// TIA Portal V19 export
FUNCTION_BLOCK "ALL_VALVES"   // FB1, LAD
{ S7_Optimized_Access := 'TRUE' }
// stored: MemoryReserve 100, SetENOAutomatically false
   VAR
      valve_R1_XV01 { S7_SetPoint := 'True'} : "valve";
      valve_R1_XV02 { S7_SetPoint := 'True'} : "valve";
      valve_R1_XV03 { S7_SetPoint := 'True'} : "valve";
      valve_R1_XV04 { S7_SetPoint := 'True'} : "valve";
      valve_R1_XV05 { S7_SetPoint := 'True'} : "valve";
      valve_R1_XV06 { S7_SetPoint := 'True'} : "valve";
      valve_R1_XV07 { S7_SetPoint := 'True'} : "valve";
      valve_R1_XV08 { S7_SetPoint := 'True'} : "valve";
      valve_R1_XV09 { S7_SetPoint := 'True'} : "valve";
      valve_R1_XV10 { S7_SetPoint := 'True'} : "valve";
      clod_skid { S7_SetPoint := 'True'} : "valve";
      valve_R2_XV01 { S7_SetPoint := 'True'} : "valve";
      valve_R2_XV02 { S7_SetPoint := 'True'} : "valve";
      valve_R2_XV03 { S7_SetPoint := 'True'} : "valve";
      valve_R2_XV04 { S7_SetPoint := 'True'} : "valve";
      valve_R2_XV05 { S7_SetPoint := 'True'} : "valve";
      valve_R2_XV06 { S7_SetPoint := 'True'} : "valve";
      valve_R2_XV07 { S7_SetPoint := 'True'} : "valve";
      valve_R2_XV08 { S7_SetPoint := 'True'} : "valve";
      valve_R2_XV09 { S7_SetPoint := 'True'} : "valve";
      valve_R2_XV10 { S7_SetPoint := 'True'} : "valve";
      valve_R3_XV01 { S7_SetPoint := 'True'} : "valve";
      valve_R3_XV02 { S7_SetPoint := 'True'} : "valve";
      valve_R3_XV03 { S7_SetPoint := 'True'} : "valve";
      valve_R3_XV04 { S7_SetPoint := 'True'} : "valve";
      valve_R3_XV05 { S7_SetPoint := 'True'} : "valve";
      valve_R3_XV06 { S7_SetPoint := 'True'} : "valve";
      valve_R3_XV07 { S7_SetPoint := 'True'} : "valve";
      valve_R3_XV08 { S7_SetPoint := 'True'} : "valve";
      valve_R3_XV09 { S7_SetPoint := 'True'} : "valve";
      valve_R3_XV10 { S7_SetPoint := 'True'} : "valve";
      valve_R4_XV02 { S7_SetPoint := 'True'} : "valve";
      valve_R4_XV01 { S7_SetPoint := 'True'} : "valve";
      valve_R4_XV03 { S7_SetPoint := 'True'} : "valve";
      valve_R4_XV04 { S7_SetPoint := 'True'} : "valve";
      valve_R4_XV05 { S7_SetPoint := 'True'} : "valve";
      valve_R4_XV06 { S7_SetPoint := 'True'} : "valve";
      valve_R4_XV07 { S7_SetPoint := 'True'} : "valve";
      valve_R4_XV08 { S7_SetPoint := 'True'} : "valve";
      valve_R4_XV09 { S7_SetPoint := 'True'} : "valve";
      valve_R4_XV10 { S7_SetPoint := 'True'} : "valve";
      valve_R8_XV2 { S7_SetPoint := 'True'} : "valve";
      valve_R8_XV3 { S7_SetPoint := 'True'} : "valve";
      valve_R8_XV4 { S7_SetPoint := 'True'} : "valve";
      valve_R8_XV5 { S7_SetPoint := 'True'} : "valve";
      valve_R8_XV05 { S7_SetPoint := 'True'} : "valve";
      valve_R8_XV06 { S7_SetPoint := 'True'} : "valve";
      valve_R8_XV07 { S7_SetPoint := 'True'} : "valve";
      valve_R8_XV08 { S7_SetPoint := 'True'} : "valve";
      valve_R8_XV09 { S7_SetPoint := 'True'} : "valve";
      valve_R8_XV10 { S7_SetPoint := 'True'} : "valve";
      valve_R6_XV01 { S7_SetPoint := 'True'} : "valve";
      valve_R6_XV02 { S7_SetPoint := 'True'} : "valve";
      valve_R6_XV03 { S7_SetPoint := 'True'} : "valve";
      valve_R6_XV04 { S7_SetPoint := 'True'} : "valve";
      valve_R6_XV05 { S7_SetPoint := 'True'} : "valve";
      valve_R6_XV06 { S7_SetPoint := 'True'} : "valve";
      valve_R6_XV07 { S7_SetPoint := 'True'} : "valve";
      valve_R6_XV08 { S7_SetPoint := 'True'} : "valve";
      valve_R6_XV09 { S7_SetPoint := 'True'} : "valve";
      valve_R6_XV10 { S7_SetPoint := 'True'} : "valve";
      valve_R7_XV01 { S7_SetPoint := 'True'} : "valve";
      valve_R7_XV02 { S7_SetPoint := 'True'} : "valve";
      valve_R7_XV03 { S7_SetPoint := 'True'} : "valve";
      valve_R7_XV04 { S7_SetPoint := 'True'} : "valve";
      valve_R7_XV05 { S7_SetPoint := 'True'} : "valve";
      valve_R7_XV06 { S7_SetPoint := 'True'} : "valve";
      valve_R7_XV07 { S7_SetPoint := 'True'} : "valve";
      valve_R7_XV08 { S7_SetPoint := 'True'} : "valve";
      valve_R7_XV09 { S7_SetPoint := 'True'} : "valve";
      valve_R7_XV10 { S7_SetPoint := 'True'} : "valve";
      valve_R8_XV01 { S7_SetPoint := 'True'} : "valve";
      valve_R8_XV02 { S7_SetPoint := 'True'} : "valve";
      valve_R8_XV03 { S7_SetPoint := 'True'} : "valve";
      valve_R8_XV04 { S7_SetPoint := 'True'} : "valve";
      valve_R5_XV2 { S7_SetPoint := 'True'} : "valve";
      valve_R5_XV3 { S7_SetPoint := 'True'} : "valve";
      valve_R5_XV4 { S7_SetPoint := 'True'} : "valve";
      valve_R5_XV5 { S7_SetPoint := 'True'} : "valve";
      valve_R5_XV05 { S7_SetPoint := 'True'} : "valve";
      valve_R5_XV06 { S7_SetPoint := 'True'} : "valve";
      valve_R5_XV07 { S7_SetPoint := 'True'} : "valve";
      valve_R5_XV08 { S7_SetPoint := 'True'} : "valve";
      valve_R5_XV09 { S7_SetPoint := 'True'} : "valve";
      valve_R5_XV10 { S7_SetPoint := 'True'} : "valve";
      valve_R9_XV01 { S7_SetPoint := 'True'} : "valve";
      valve_R9_XV02 { S7_SetPoint := 'True'} : "valve";
      valve_R9_XV03 { S7_SetPoint := 'True'} : "valve";
      valve_R9_XV04 { S7_SetPoint := 'True'} : "valve";
      valve_R9_XV05 { S7_SetPoint := 'True'} : "valve";
      valve_R9_XV06 { S7_SetPoint := 'True'} : "valve";
      valve_R9_XV07 { S7_SetPoint := 'True'} : "valve";
      valve_R9_XV08 { S7_SetPoint := 'True'} : "valve";
      valve_R9_XV09 { S7_SetPoint := 'True'} : "valve";
      valve_R9_XV10 { S7_SetPoint := 'True'} : "valve";
      valve_R10_XV01 { S7_SetPoint := 'True'} : "valve";
      valve_R10_XV02 { S7_SetPoint := 'True'} : "valve";
      valve_R10_XV03 { S7_SetPoint := 'True'} : "valve";
      valve_R10_XV04 { S7_SetPoint := 'True'} : "valve";
      valve_R10_XV05 { S7_SetPoint := 'True'} : "valve";
      valve_R10_XV06 { S7_SetPoint := 'True'} : "valve";
      valve_R10_XV07 { S7_SetPoint := 'True'} : "valve";
      valve_R10_XV08 { S7_SetPoint := 'True'} : "valve";
      valve_R10_XV09 { S7_SetPoint := 'True'} : "valve";
      valve_R10_XV10 { S7_SetPoint := 'True'} : "valve";
      valve_R11_XV01 { S7_SetPoint := 'True'} : "valve";
      valve_R11_XV02 { S7_SetPoint := 'True'} : "valve";
      valve_R11_XV03 { S7_SetPoint := 'True'} : "valve";
      valve_R11_XV04 { S7_SetPoint := 'True'} : "valve";
      valve_R11_XV05 { S7_SetPoint := 'True'} : "valve";
      valve_R11_XV06 { S7_SetPoint := 'True'} : "valve";
      valve_R11_XV07 { S7_SetPoint := 'True'} : "valve";
      valve_R11_XV08 { S7_SetPoint := 'True'} : "valve";
      valve_R11_XV09 { S7_SetPoint := 'True'} : "valve";
      valve_R11_XV10 { S7_SetPoint := 'True'} : "valve";
      valve_R12_XV01 { S7_SetPoint := 'True'} : "valve";
      valve_R12_XV02 { S7_SetPoint := 'True'} : "valve";
      valve_R12_XV03 { S7_SetPoint := 'True'} : "valve";
      valve_R12_XV04 { S7_SetPoint := 'True'} : "valve";
      valve_R12_XV05 { S7_SetPoint := 'True'} : "valve";
      valve_R12_XV06 { S7_SetPoint := 'True'} : "valve";
      valve_R12_XV07 { S7_SetPoint := 'True'} : "valve";
      valve_R12_XV08 { S7_SetPoint := 'True'} : "valve";
      valve_R12_XV09 { S7_SetPoint := 'True'} : "valve";
      valve_R12_XV10 { S7_SetPoint := 'True'} : "valve";
      valve_R13_XV01 { S7_SetPoint := 'True'} : "valve";
      valve_R13_XV02 { S7_SetPoint := 'True'} : "valve";
      valve_R13_XV03 { S7_SetPoint := 'True'} : "valve";
      valve_R13_XV04 { S7_SetPoint := 'True'} : "valve";
      valve_R13_XV05 { S7_SetPoint := 'True'} : "valve";
      valve_R13_XV06 { S7_SetPoint := 'True'} : "valve";
      valve_R13_XV07 { S7_SetPoint := 'True'} : "valve";
      valve_R13_XV08 { S7_SetPoint := 'True'} : "valve";
      valve_R13_XV09 { S7_SetPoint := 'True'} : "valve";
      valve_R13_XV10 { S7_SetPoint := 'True'} : "valve";
      valve_R14_XV02 { S7_SetPoint := 'True'} : "valve";
      valve_R14_XV01 { S7_SetPoint := 'True'} : "valve";
      valve_R14_XV03 { S7_SetPoint := 'True'} : "valve";
      valve_R14_XV04 { S7_SetPoint := 'True'} : "valve";
      valve_R14_XV05 { S7_SetPoint := 'True'} : "valve";
      valve_R14_XV06 { S7_SetPoint := 'True'} : "valve";
      valve_R14_XV07 { S7_SetPoint := 'True'} : "valve";
      valve_R14_XV08 { S7_SetPoint := 'True'} : "valve";
      valve_R14_XV09 { S7_SetPoint := 'True'} : "valve";
      valve_R14_XV10 { S7_SetPoint := 'True'} : "valve";
      valve_R15_XV02 { S7_SetPoint := 'True'} : "valve";
      valve_R15_XV01 { S7_SetPoint := 'True'} : "valve";
      valve_R15_XV03 { S7_SetPoint := 'True'} : "valve";
      valve_R15_XV04 { S7_SetPoint := 'True'} : "valve";
      valve_R15_XV05 { S7_SetPoint := 'True'} : "valve";
      valve_R15_XV06 { S7_SetPoint := 'True'} : "valve";
      valve_R15_XV07 { S7_SetPoint := 'True'} : "valve";
      valve_R15_XV08 { S7_SetPoint := 'True'} : "valve";
      valve_R15_XV09 { S7_SetPoint := 'True'} : "valve";
      valve_R15_XV10 { S7_SetPoint := 'True'} : "valve";
      valve_R16_XV02 { S7_SetPoint := 'True'} : "valve";
      valve_R16_XV03 { S7_SetPoint := 'True'} : "valve";
      valve_R16_XV04 { S7_SetPoint := 'True'} : "valve";
      valve_R16_XV05 { S7_SetPoint := 'True'} : "valve";
      valve_R16_XV06 { S7_SetPoint := 'True'} : "valve";
      valve_R16_XV07 { S7_SetPoint := 'True'} : "valve";
      valve_R16_XV08 { S7_SetPoint := 'True'} : "valve";
      valve_R16_XV09 { S7_SetPoint := 'True'} : "valve";
      valve_R16_XV10 { S7_SetPoint := 'True'} : "valve";
      valve_R17_XV01 { S7_SetPoint := 'True'} : "valve";
      valve_R17_XV02 { S7_SetPoint := 'True'} : "valve";
      valve_R17_XV03 { S7_SetPoint := 'True'} : "valve";
      valve_R17_XV04 { S7_SetPoint := 'True'} : "valve";
      valve_R17_XV05 { S7_SetPoint := 'True'} : "valve";
      valve_R17_XV06 { S7_SetPoint := 'True'} : "valve";
      valve_R17_XV07 { S7_SetPoint := 'True'} : "valve";
      valve_R17_XV08 { S7_SetPoint := 'True'} : "valve";
      valve_R17_XV09 { S7_SetPoint := 'True'} : "valve";
      valve_R17_XV10 { S7_SetPoint := 'True'} : "valve";
      valve_R18_XV02 { S7_SetPoint := 'True'} : "valve";
      valve_R18_XV03 { S7_SetPoint := 'True'} : "valve";
      valve_R18_XV04 { S7_SetPoint := 'True'} : "valve";
      valve_R18_XV05 { S7_SetPoint := 'True'} : "valve";
      valve_R18_XV06 { S7_SetPoint := 'True'} : "valve";
      valve_R18_XV07 { S7_SetPoint := 'True'} : "valve";
      valve_R18_XV08 { S7_SetPoint := 'True'} : "valve";
      valve_R18_XV09 { S7_SetPoint := 'True'} : "valve";
      valve_R18_XV10 { S7_SetPoint := 'True'} : "valve";
      child_skid { S7_SetPoint := 'True'} : "valve";
      ultra_child { S7_SetPoint := 'True'} : "valve";
   END_VAR
BEGIN

REGION Network 1: R1_XV01
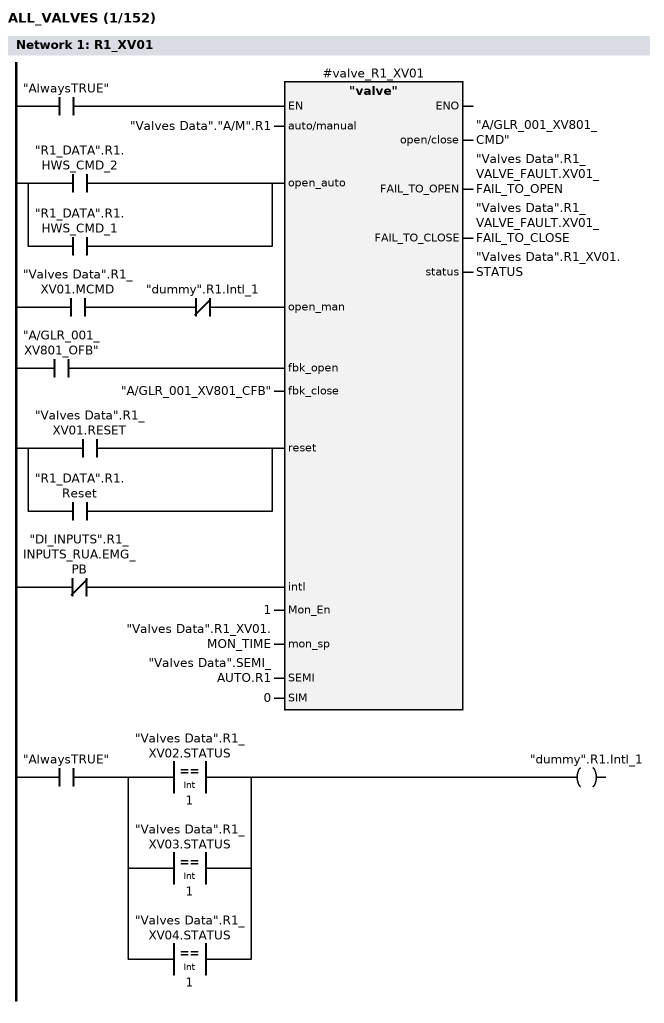
   RUNG wire#powerrail
      Contact( "AlwaysTRUE" )
      #valve_R1_XV01(open_auto := wire#w1, open_man := wire#w2, fbk_open := wire#w3, reset := wire#w4, intl := wire#w5, "auto/manual" := "Valves Data"."A/M".R1, fbk_close := "A/GLR_001_XV801_CFB", Mon_En := 1, mon_sp := "Valves Data".R1_XV01.MON_TIME, SEMI := "Valves Data".SEMI_AUTO.R1, SIM := 0, "open/close" => "A/GLR_001_XV801_CMD", FAIL_TO_OPEN => "Valves Data".R1_VALVE_FAULT.XV01_FAIL_TO_OPEN, FAIL_TO_CLOSE => "Valves Data".R1_VALVE_FAULT.XV01_FAIL_TO_CLOSE, status => "Valves Data".R1_XV01.STATUS)
   END_RUNG
   RUNG wire#powerrail
      Contact( "R1_DATA".R1.HWS_CMD_2 )
   END_RUNG wire#w1
   RUNG wire#powerrail
      Contact( "R1_DATA".R1.HWS_CMD_1 )
   END_RUNG wire#w1
   RUNG wire#powerrail
      Contact( "Valves Data".R1_XV01.MCMD )
      I_Contact( "dummy".R1.Intl_1 )
   END_RUNG wire#w2
   RUNG wire#powerrail
      Contact( "A/GLR_001_XV801_OFB" )
   END_RUNG wire#w3
   RUNG wire#powerrail
      Contact( "Valves Data".R1_XV01.RESET )
   END_RUNG wire#w4
   RUNG wire#powerrail
      Contact( "R1_DATA".R1.Reset )
   END_RUNG wire#w4
   RUNG wire#powerrail
      I_Contact( "DI_INPUTS".R1_INPUTS_RUA.EMG_PB )
   END_RUNG wire#w5
   RUNG wire#powerrail
      Contact( "AlwaysTRUE" )
      wire#w6
      { S7_Templates := "SrcType := Int" } EQ_Contact(in1 := "Valves Data".R1_XV02.STATUS, in2 := 1)
      wire#w7
      Coil( "dummy".R1.Intl_1 )
   END_RUNG
   RUNG wire#w6
      { S7_Templates := "SrcType := Int" } EQ_Contact(in1 := "Valves Data".R1_XV03.STATUS, in2 := 1)
   END_RUNG wire#w7
   RUNG wire#w6
      { S7_Templates := "SrcType := Int" } EQ_Contact(in1 := "Valves Data".R1_XV04.STATUS, in2 := 1)
   END_RUNG wire#w7
   // the same network as SCL:
   IF "AlwaysTRUE" THEN
       #valve_R1_XV01("auto/manual" := "Valves Data"."A/M".R1,   // "valve"
                      open_auto := "R1_DATA".R1.HWS_CMD_2 OR "R1_DATA".R1.HWS_CMD_1,
                      open_man := "Valves Data".R1_XV01.MCMD AND NOT "dummy".R1.Intl_1,
                      fbk_open := "A/GLR_001_XV801_OFB",
                      fbk_close := "A/GLR_001_XV801_CFB",
                      reset := "Valves Data".R1_XV01.RESET OR "R1_DATA".R1.Reset,
                      intl := NOT "DI_INPUTS".R1_INPUTS_RUA.EMG_PB,
                      Mon_En := 1,
                      mon_sp := "Valves Data".R1_XV01.MON_TIME,
                      SEMI := "Valves Data".SEMI_AUTO.R1,
                      SIM := 0,
                      "open/close" => "A/GLR_001_XV801_CMD",
                      FAIL_TO_OPEN => "Valves Data".R1_VALVE_FAULT.XV01_FAIL_TO_OPEN,
                      FAIL_TO_CLOSE => "Valves Data".R1_VALVE_FAULT.XV01_FAIL_TO_CLOSE,
                      status => "Valves Data".R1_XV01.STATUS);
   END_IF;
   "dummy".R1.Intl_1 := "AlwaysTRUE" AND (("Valves Data".R1_XV02.STATUS = 1) OR ("Valves Data".R1_XV03.STATUS = 1) OR ("Valves Data".R1_XV04.STATUS = 1));
END_REGION

REGION Network 2: R1_XV02
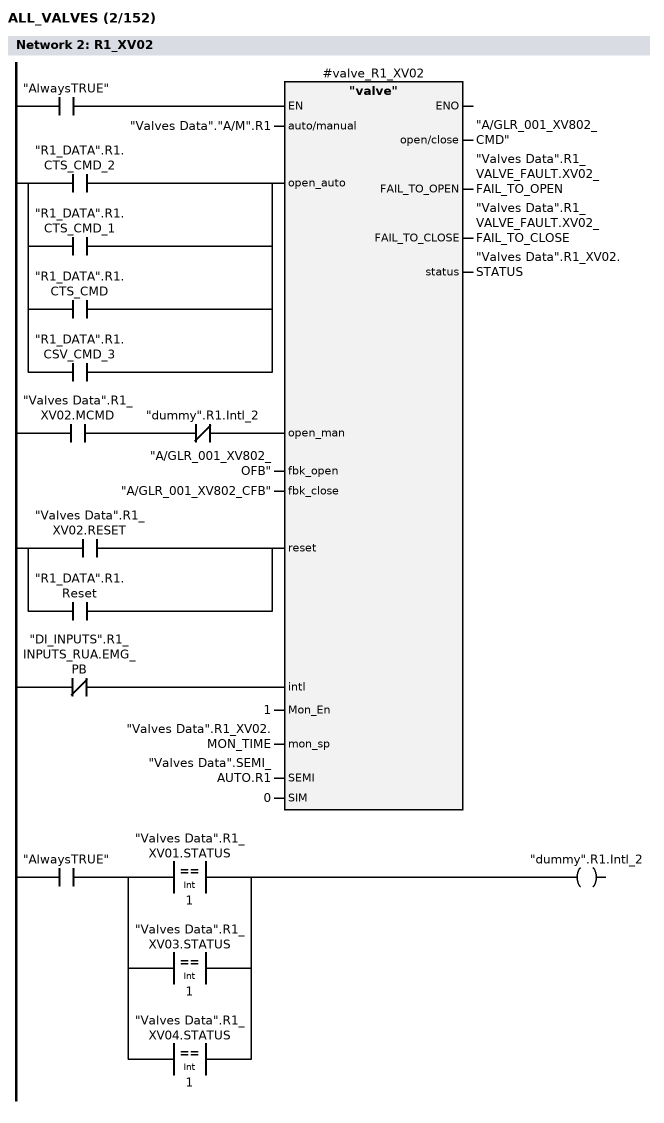
   RUNG wire#powerrail
      Contact( "AlwaysTRUE" )
      #valve_R1_XV02(open_auto := wire#w1, open_man := wire#w2, reset := wire#w3, intl := wire#w4, "auto/manual" := "Valves Data"."A/M".R1, fbk_open := "A/GLR_001_XV802_OFB", fbk_close := "A/GLR_001_XV802_CFB", Mon_En := 1, mon_sp := "Valves Data".R1_XV02.MON_TIME, SEMI := "Valves Data".SEMI_AUTO.R1, SIM := 0, "open/close" => "A/GLR_001_XV802_CMD", FAIL_TO_OPEN => "Valves Data".R1_VALVE_FAULT.XV02_FAIL_TO_OPEN, FAIL_TO_CLOSE => "Valves Data".R1_VALVE_FAULT.XV02_FAIL_TO_CLOSE, status => "Valves Data".R1_XV02.STATUS)
   END_RUNG
   RUNG wire#powerrail
      Contact( "R1_DATA".R1.CTS_CMD_2 )
   END_RUNG wire#w1
   RUNG wire#powerrail
      Contact( "R1_DATA".R1.CTS_CMD_1 )
   END_RUNG wire#w1
   RUNG wire#powerrail
      Contact( "R1_DATA".R1.CTS_CMD )
   END_RUNG wire#w1
   RUNG wire#powerrail
      Contact( "R1_DATA".R1.CSV_CMD_3 )
   END_RUNG wire#w1
   RUNG wire#powerrail
      Contact( "Valves Data".R1_XV02.MCMD )
      I_Contact( "dummy".R1.Intl_2 )
   END_RUNG wire#w2
   RUNG wire#powerrail
      Contact( "Valves Data".R1_XV02.RESET )
   END_RUNG wire#w3
   RUNG wire#powerrail
      Contact( "R1_DATA".R1.Reset )
   END_RUNG wire#w3
   RUNG wire#powerrail
      I_Contact( "DI_INPUTS".R1_INPUTS_RUA.EMG_PB )
   END_RUNG wire#w4
   RUNG wire#powerrail
      Contact( "AlwaysTRUE" )
      wire#w5
      { S7_Templates := "SrcType := Int" } EQ_Contact(in1 := "Valves Data".R1_XV01.STATUS, in2 := 1)
      wire#w6
      Coil( "dummy".R1.Intl_2 )
   END_RUNG
   RUNG wire#w5
      { S7_Templates := "SrcType := Int" } EQ_Contact(in1 := "Valves Data".R1_XV03.STATUS, in2 := 1)
   END_RUNG wire#w6
   RUNG wire#w5
      { S7_Templates := "SrcType := Int" } EQ_Contact(in1 := "Valves Data".R1_XV04.STATUS, in2 := 1)
   END_RUNG wire#w6
   // the same network as SCL:
   IF "AlwaysTRUE" THEN
       #valve_R1_XV02("auto/manual" := "Valves Data"."A/M".R1,   // "valve"
                      open_auto := "R1_DATA".R1.CTS_CMD_2 OR "R1_DATA".R1.CTS_CMD_1 OR "R1_DATA".R1.CTS_CMD OR "R1_DATA".R1.CSV_CMD_3,
                      open_man := "Valves Data".R1_XV02.MCMD AND NOT "dummy".R1.Intl_2,
                      fbk_open := "A/GLR_001_XV802_OFB",
                      fbk_close := "A/GLR_001_XV802_CFB",
                      reset := "Valves Data".R1_XV02.RESET OR "R1_DATA".R1.Reset,
                      intl := NOT "DI_INPUTS".R1_INPUTS_RUA.EMG_PB,
                      Mon_En := 1,
                      mon_sp := "Valves Data".R1_XV02.MON_TIME,
                      SEMI := "Valves Data".SEMI_AUTO.R1,
                      SIM := 0,
                      "open/close" => "A/GLR_001_XV802_CMD",
                      FAIL_TO_OPEN => "Valves Data".R1_VALVE_FAULT.XV02_FAIL_TO_OPEN,
                      FAIL_TO_CLOSE => "Valves Data".R1_VALVE_FAULT.XV02_FAIL_TO_CLOSE,
                      status => "Valves Data".R1_XV02.STATUS);
   END_IF;
   "dummy".R1.Intl_2 := "AlwaysTRUE" AND (("Valves Data".R1_XV01.STATUS = 1) OR ("Valves Data".R1_XV03.STATUS = 1) OR ("Valves Data".R1_XV04.STATUS = 1));
END_REGION

REGION Network 3: R1_XV03
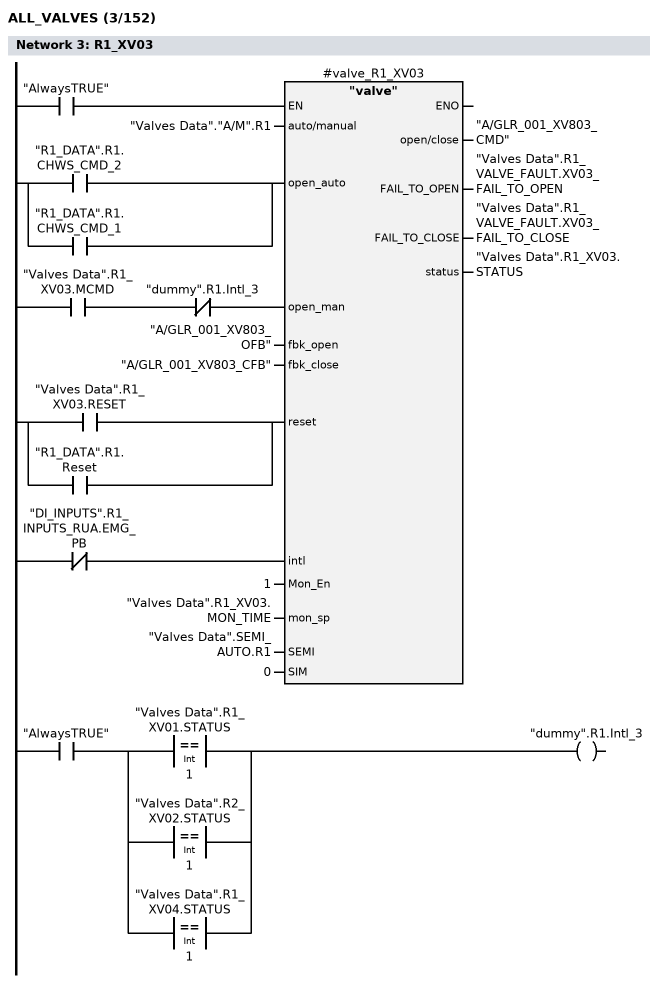
   RUNG wire#powerrail
      Contact( "AlwaysTRUE" )
      #valve_R1_XV03(open_auto := wire#w1, open_man := wire#w2, reset := wire#w3, intl := wire#w4, "auto/manual" := "Valves Data"."A/M".R1, fbk_open := "A/GLR_001_XV803_OFB", fbk_close := "A/GLR_001_XV803_CFB", Mon_En := 1, mon_sp := "Valves Data".R1_XV03.MON_TIME, SEMI := "Valves Data".SEMI_AUTO.R1, SIM := 0, "open/close" => "A/GLR_001_XV803_CMD", FAIL_TO_OPEN => "Valves Data".R1_VALVE_FAULT.XV03_FAIL_TO_OPEN, FAIL_TO_CLOSE => "Valves Data".R1_VALVE_FAULT.XV03_FAIL_TO_CLOSE, status => "Valves Data".R1_XV03.STATUS)
   END_RUNG
   RUNG wire#powerrail
      Contact( "R1_DATA".R1.CHWS_CMD_2 )
   END_RUNG wire#w1
   RUNG wire#powerrail
      Contact( "R1_DATA".R1.CHWS_CMD_1 )
   END_RUNG wire#w1
   RUNG wire#powerrail
      Contact( "Valves Data".R1_XV03.MCMD )
      I_Contact( "dummy".R1.Intl_3 )
   END_RUNG wire#w2
   RUNG wire#powerrail
      Contact( "Valves Data".R1_XV03.RESET )
   END_RUNG wire#w3
   RUNG wire#powerrail
      Contact( "R1_DATA".R1.Reset )
   END_RUNG wire#w3
   RUNG wire#powerrail
      I_Contact( "DI_INPUTS".R1_INPUTS_RUA.EMG_PB )
   END_RUNG wire#w4
   RUNG wire#powerrail
      Contact( "AlwaysTRUE" )
      wire#w5
      { S7_Templates := "SrcType := Int" } EQ_Contact(in1 := "Valves Data".R1_XV01.STATUS, in2 := 1)
      wire#w6
      Coil( "dummy".R1.Intl_3 )
   END_RUNG
   RUNG wire#w5
      { S7_Templates := "SrcType := Int" } EQ_Contact(in1 := "Valves Data".R2_XV02.STATUS, in2 := 1)
   END_RUNG wire#w6
   RUNG wire#w5
      { S7_Templates := "SrcType := Int" } EQ_Contact(in1 := "Valves Data".R1_XV04.STATUS, in2 := 1)
   END_RUNG wire#w6
   // the same network as SCL:
   IF "AlwaysTRUE" THEN
       #valve_R1_XV03("auto/manual" := "Valves Data"."A/M".R1,   // "valve"
                      open_auto := "R1_DATA".R1.CHWS_CMD_2 OR "R1_DATA".R1.CHWS_CMD_1,
                      open_man := "Valves Data".R1_XV03.MCMD AND NOT "dummy".R1.Intl_3,
                      fbk_open := "A/GLR_001_XV803_OFB",
                      fbk_close := "A/GLR_001_XV803_CFB",
                      reset := "Valves Data".R1_XV03.RESET OR "R1_DATA".R1.Reset,
                      intl := NOT "DI_INPUTS".R1_INPUTS_RUA.EMG_PB,
                      Mon_En := 1,
                      mon_sp := "Valves Data".R1_XV03.MON_TIME,
                      SEMI := "Valves Data".SEMI_AUTO.R1,
                      SIM := 0,
                      "open/close" => "A/GLR_001_XV803_CMD",
                      FAIL_TO_OPEN => "Valves Data".R1_VALVE_FAULT.XV03_FAIL_TO_OPEN,
                      FAIL_TO_CLOSE => "Valves Data".R1_VALVE_FAULT.XV03_FAIL_TO_CLOSE,
                      status => "Valves Data".R1_XV03.STATUS);
   END_IF;
   "dummy".R1.Intl_3 := "AlwaysTRUE" AND (("Valves Data".R1_XV01.STATUS = 1) OR ("Valves Data".R2_XV02.STATUS = 1) OR ("Valves Data".R1_XV04.STATUS = 1));
END_REGION

REGION Network 4: R1_XV04
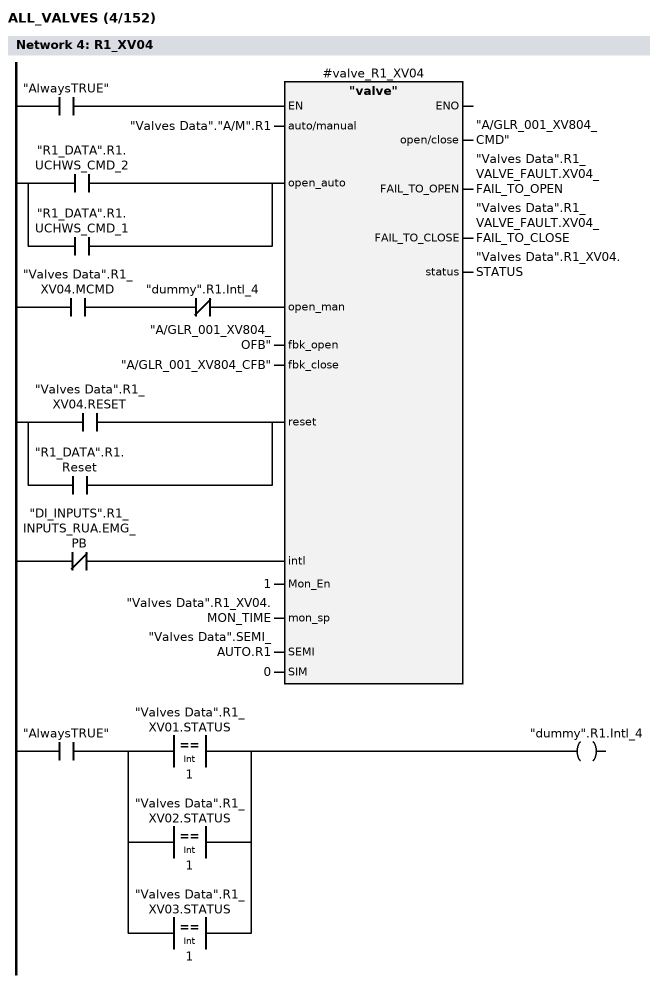
   RUNG wire#powerrail
      Contact( "AlwaysTRUE" )
      #valve_R1_XV04(open_auto := wire#w1, open_man := wire#w2, reset := wire#w3, intl := wire#w4, "auto/manual" := "Valves Data"."A/M".R1, fbk_open := "A/GLR_001_XV804_OFB", fbk_close := "A/GLR_001_XV804_CFB", Mon_En := 1, mon_sp := "Valves Data".R1_XV04.MON_TIME, SEMI := "Valves Data".SEMI_AUTO.R1, SIM := 0, "open/close" => "A/GLR_001_XV804_CMD", FAIL_TO_OPEN => "Valves Data".R1_VALVE_FAULT.XV04_FAIL_TO_OPEN, FAIL_TO_CLOSE => "Valves Data".R1_VALVE_FAULT.XV04_FAIL_TO_CLOSE, status => "Valves Data".R1_XV04.STATUS)
   END_RUNG
   RUNG wire#powerrail
      Contact( "R1_DATA".R1.UCHWS_CMD_2 )
   END_RUNG wire#w1
   RUNG wire#powerrail
      Contact( "R1_DATA".R1.UCHWS_CMD_1 )
   END_RUNG wire#w1
   RUNG wire#powerrail
      Contact( "Valves Data".R1_XV04.MCMD )
      I_Contact( "dummy".R1.Intl_4 )
   END_RUNG wire#w2
   RUNG wire#powerrail
      Contact( "Valves Data".R1_XV04.RESET )
   END_RUNG wire#w3
   RUNG wire#powerrail
      Contact( "R1_DATA".R1.Reset )
   END_RUNG wire#w3
   RUNG wire#powerrail
      I_Contact( "DI_INPUTS".R1_INPUTS_RUA.EMG_PB )
   END_RUNG wire#w4
   RUNG wire#powerrail
      Contact( "AlwaysTRUE" )
      wire#w5
      { S7_Templates := "SrcType := Int" } EQ_Contact(in1 := "Valves Data".R1_XV01.STATUS, in2 := 1)
      wire#w6
      Coil( "dummy".R1.Intl_4 )
   END_RUNG
   RUNG wire#w5
      { S7_Templates := "SrcType := Int" } EQ_Contact(in1 := "Valves Data".R1_XV02.STATUS, in2 := 1)
   END_RUNG wire#w6
   RUNG wire#w5
      { S7_Templates := "SrcType := Int" } EQ_Contact(in1 := "Valves Data".R1_XV03.STATUS, in2 := 1)
   END_RUNG wire#w6
   // the same network as SCL:
   IF "AlwaysTRUE" THEN
       #valve_R1_XV04("auto/manual" := "Valves Data"."A/M".R1,   // "valve"
                      open_auto := "R1_DATA".R1.UCHWS_CMD_2 OR "R1_DATA".R1.UCHWS_CMD_1,
                      open_man := "Valves Data".R1_XV04.MCMD AND NOT "dummy".R1.Intl_4,
                      fbk_open := "A/GLR_001_XV804_OFB",
                      fbk_close := "A/GLR_001_XV804_CFB",
                      reset := "Valves Data".R1_XV04.RESET OR "R1_DATA".R1.Reset,
                      intl := NOT "DI_INPUTS".R1_INPUTS_RUA.EMG_PB,
                      Mon_En := 1,
                      mon_sp := "Valves Data".R1_XV04.MON_TIME,
                      SEMI := "Valves Data".SEMI_AUTO.R1,
                      SIM := 0,
                      "open/close" => "A/GLR_001_XV804_CMD",
                      FAIL_TO_OPEN => "Valves Data".R1_VALVE_FAULT.XV04_FAIL_TO_OPEN,
                      FAIL_TO_CLOSE => "Valves Data".R1_VALVE_FAULT.XV04_FAIL_TO_CLOSE,
                      status => "Valves Data".R1_XV04.STATUS);
   END_IF;
   "dummy".R1.Intl_4 := "AlwaysTRUE" AND (("Valves Data".R1_XV01.STATUS = 1) OR ("Valves Data".R1_XV02.STATUS = 1) OR ("Valves Data".R1_XV03.STATUS = 1));
END_REGION

REGION Network 5: R1_XV05
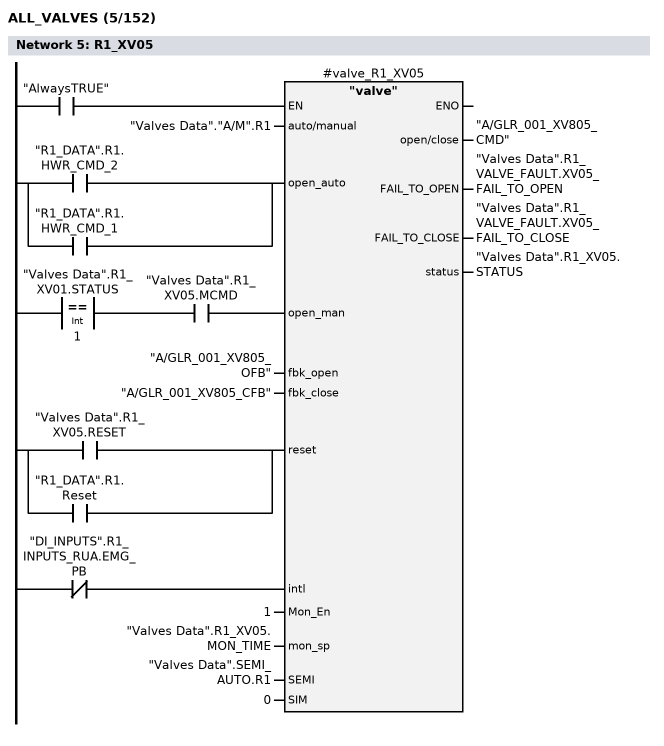
   RUNG wire#powerrail
      Contact( "AlwaysTRUE" )
      #valve_R1_XV05(open_auto := wire#w1, open_man := wire#w2, reset := wire#w3, intl := wire#w4, "auto/manual" := "Valves Data"."A/M".R1, fbk_open := "A/GLR_001_XV805_OFB", fbk_close := "A/GLR_001_XV805_CFB", Mon_En := 1, mon_sp := "Valves Data".R1_XV05.MON_TIME, SEMI := "Valves Data".SEMI_AUTO.R1, SIM := 0, "open/close" => "A/GLR_001_XV805_CMD", FAIL_TO_OPEN => "Valves Data".R1_VALVE_FAULT.XV05_FAIL_TO_OPEN, FAIL_TO_CLOSE => "Valves Data".R1_VALVE_FAULT.XV05_FAIL_TO_CLOSE, status => "Valves Data".R1_XV05.STATUS)
   END_RUNG
   RUNG wire#powerrail
      Contact( "R1_DATA".R1.HWR_CMD_2 )
   END_RUNG wire#w1
   RUNG wire#powerrail
      Contact( "R1_DATA".R1.HWR_CMD_1 )
   END_RUNG wire#w1
   RUNG wire#powerrail
      { S7_Templates := "SrcType := Int" } EQ_Contact(in1 := "Valves Data".R1_XV01.STATUS, in2 := 1)
      Contact( "Valves Data".R1_XV05.MCMD )
   END_RUNG wire#w2
   RUNG wire#powerrail
      Contact( "Valves Data".R1_XV05.RESET )
   END_RUNG wire#w3
   RUNG wire#powerrail
      Contact( "R1_DATA".R1.Reset )
   END_RUNG wire#w3
   RUNG wire#powerrail
      I_Contact( "DI_INPUTS".R1_INPUTS_RUA.EMG_PB )
   END_RUNG wire#w4
   // the same network as SCL:
   IF "AlwaysTRUE" THEN
       #valve_R1_XV05("auto/manual" := "Valves Data"."A/M".R1,   // "valve"
                      open_auto := "R1_DATA".R1.HWR_CMD_2 OR "R1_DATA".R1.HWR_CMD_1,
                      open_man := ("Valves Data".R1_XV01.STATUS = 1) AND "Valves Data".R1_XV05.MCMD,
                      fbk_open := "A/GLR_001_XV805_OFB",
                      fbk_close := "A/GLR_001_XV805_CFB",
                      reset := "Valves Data".R1_XV05.RESET OR "R1_DATA".R1.Reset,
                      intl := NOT "DI_INPUTS".R1_INPUTS_RUA.EMG_PB,
                      Mon_En := 1,
                      mon_sp := "Valves Data".R1_XV05.MON_TIME,
                      SEMI := "Valves Data".SEMI_AUTO.R1,
                      SIM := 0,
                      "open/close" => "A/GLR_001_XV805_CMD",
                      FAIL_TO_OPEN => "Valves Data".R1_VALVE_FAULT.XV05_FAIL_TO_OPEN,
                      FAIL_TO_CLOSE => "Valves Data".R1_VALVE_FAULT.XV05_FAIL_TO_CLOSE,
                      status => "Valves Data".R1_XV05.STATUS);
   END_IF;
END_REGION

REGION Network 6: R1_XV06
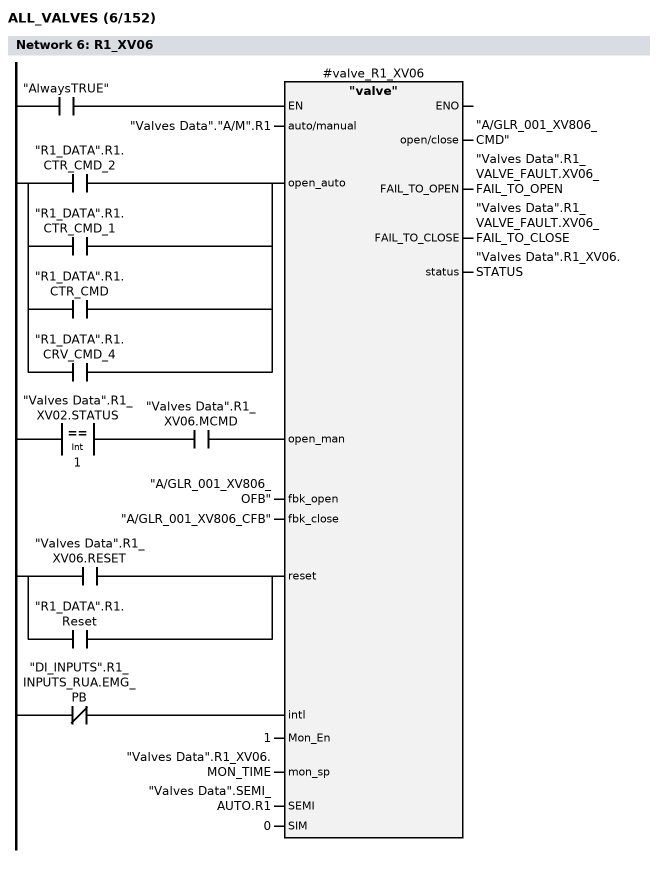
   RUNG wire#powerrail
      Contact( "AlwaysTRUE" )
      #valve_R1_XV06(open_auto := wire#w1, open_man := wire#w2, reset := wire#w3, intl := wire#w4, "auto/manual" := "Valves Data"."A/M".R1, fbk_open := "A/GLR_001_XV806_OFB", fbk_close := "A/GLR_001_XV806_CFB", Mon_En := 1, mon_sp := "Valves Data".R1_XV06.MON_TIME, SEMI := "Valves Data".SEMI_AUTO.R1, SIM := 0, "open/close" => "A/GLR_001_XV806_CMD", FAIL_TO_OPEN => "Valves Data".R1_VALVE_FAULT.XV06_FAIL_TO_OPEN, FAIL_TO_CLOSE => "Valves Data".R1_VALVE_FAULT.XV06_FAIL_TO_CLOSE, status => "Valves Data".R1_XV06.STATUS)
   END_RUNG
   RUNG wire#powerrail
      Contact( "R1_DATA".R1.CTR_CMD_2 )
   END_RUNG wire#w1
   RUNG wire#powerrail
      Contact( "R1_DATA".R1.CTR_CMD_1 )
   END_RUNG wire#w1
   RUNG wire#powerrail
      Contact( "R1_DATA".R1.CTR_CMD )
   END_RUNG wire#w1
   RUNG wire#powerrail
      Contact( "R1_DATA".R1.CRV_CMD_4 )
   END_RUNG wire#w1
   RUNG wire#powerrail
      { S7_Templates := "SrcType := Int" } EQ_Contact(in1 := "Valves Data".R1_XV02.STATUS, in2 := 1)
      Contact( "Valves Data".R1_XV06.MCMD )
   END_RUNG wire#w2
   RUNG wire#powerrail
      Contact( "Valves Data".R1_XV06.RESET )
   END_RUNG wire#w3
   RUNG wire#powerrail
      Contact( "R1_DATA".R1.Reset )
   END_RUNG wire#w3
   RUNG wire#powerrail
      I_Contact( "DI_INPUTS".R1_INPUTS_RUA.EMG_PB )
   END_RUNG wire#w4
   // the same network as SCL:
   IF "AlwaysTRUE" THEN
       #valve_R1_XV06("auto/manual" := "Valves Data"."A/M".R1,   // "valve"
                      open_auto := "R1_DATA".R1.CTR_CMD_2 OR "R1_DATA".R1.CTR_CMD_1 OR "R1_DATA".R1.CTR_CMD OR "R1_DATA".R1.CRV_CMD_4,
                      open_man := ("Valves Data".R1_XV02.STATUS = 1) AND "Valves Data".R1_XV06.MCMD,
                      fbk_open := "A/GLR_001_XV806_OFB",
                      fbk_close := "A/GLR_001_XV806_CFB",
                      reset := "Valves Data".R1_XV06.RESET OR "R1_DATA".R1.Reset,
                      intl := NOT "DI_INPUTS".R1_INPUTS_RUA.EMG_PB,
                      Mon_En := 1,
                      mon_sp := "Valves Data".R1_XV06.MON_TIME,
                      SEMI := "Valves Data".SEMI_AUTO.R1,
                      SIM := 0,
                      "open/close" => "A/GLR_001_XV806_CMD",
                      FAIL_TO_OPEN => "Valves Data".R1_VALVE_FAULT.XV06_FAIL_TO_OPEN,
                      FAIL_TO_CLOSE => "Valves Data".R1_VALVE_FAULT.XV06_FAIL_TO_CLOSE,
                      status => "Valves Data".R1_XV06.STATUS);
   END_IF;
END_REGION

REGION Network 7: R1_XV07
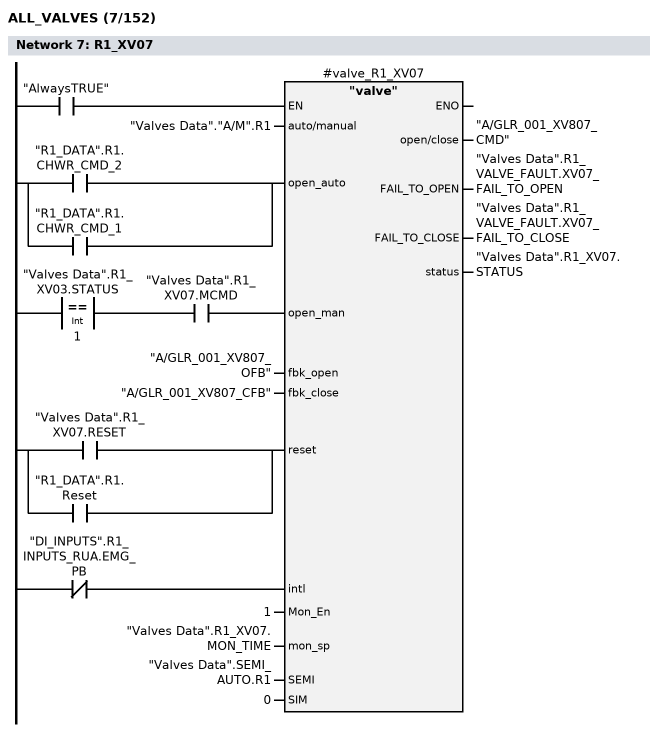
   RUNG wire#powerrail
      Contact( "AlwaysTRUE" )
      #valve_R1_XV07(open_auto := wire#w1, open_man := wire#w2, reset := wire#w3, intl := wire#w4, "auto/manual" := "Valves Data"."A/M".R1, fbk_open := "A/GLR_001_XV807_OFB", fbk_close := "A/GLR_001_XV807_CFB", Mon_En := 1, mon_sp := "Valves Data".R1_XV07.MON_TIME, SEMI := "Valves Data".SEMI_AUTO.R1, SIM := 0, "open/close" => "A/GLR_001_XV807_CMD", FAIL_TO_OPEN => "Valves Data".R1_VALVE_FAULT.XV07_FAIL_TO_OPEN, FAIL_TO_CLOSE => "Valves Data".R1_VALVE_FAULT.XV07_FAIL_TO_CLOSE, status => "Valves Data".R1_XV07.STATUS)
   END_RUNG
   RUNG wire#powerrail
      Contact( "R1_DATA".R1.CHWR_CMD_2 )
   END_RUNG wire#w1
   RUNG wire#powerrail
      Contact( "R1_DATA".R1.CHWR_CMD_1 )
   END_RUNG wire#w1
   RUNG wire#powerrail
      { S7_Templates := "SrcType := Int" } EQ_Contact(in1 := "Valves Data".R1_XV03.STATUS, in2 := 1)
      Contact( "Valves Data".R1_XV07.MCMD )
   END_RUNG wire#w2
   RUNG wire#powerrail
      Contact( "Valves Data".R1_XV07.RESET )
   END_RUNG wire#w3
   RUNG wire#powerrail
      Contact( "R1_DATA".R1.Reset )
   END_RUNG wire#w3
   RUNG wire#powerrail
      I_Contact( "DI_INPUTS".R1_INPUTS_RUA.EMG_PB )
   END_RUNG wire#w4
   // the same network as SCL:
   IF "AlwaysTRUE" THEN
       #valve_R1_XV07("auto/manual" := "Valves Data"."A/M".R1,   // "valve"
                      open_auto := "R1_DATA".R1.CHWR_CMD_2 OR "R1_DATA".R1.CHWR_CMD_1,
                      open_man := ("Valves Data".R1_XV03.STATUS = 1) AND "Valves Data".R1_XV07.MCMD,
                      fbk_open := "A/GLR_001_XV807_OFB",
                      fbk_close := "A/GLR_001_XV807_CFB",
                      reset := "Valves Data".R1_XV07.RESET OR "R1_DATA".R1.Reset,
                      intl := NOT "DI_INPUTS".R1_INPUTS_RUA.EMG_PB,
                      Mon_En := 1,
                      mon_sp := "Valves Data".R1_XV07.MON_TIME,
                      SEMI := "Valves Data".SEMI_AUTO.R1,
                      SIM := 0,
                      "open/close" => "A/GLR_001_XV807_CMD",
                      FAIL_TO_OPEN => "Valves Data".R1_VALVE_FAULT.XV07_FAIL_TO_OPEN,
                      FAIL_TO_CLOSE => "Valves Data".R1_VALVE_FAULT.XV07_FAIL_TO_CLOSE,
                      status => "Valves Data".R1_XV07.STATUS);
   END_IF;
END_REGION

REGION Network 8: R1_XV08
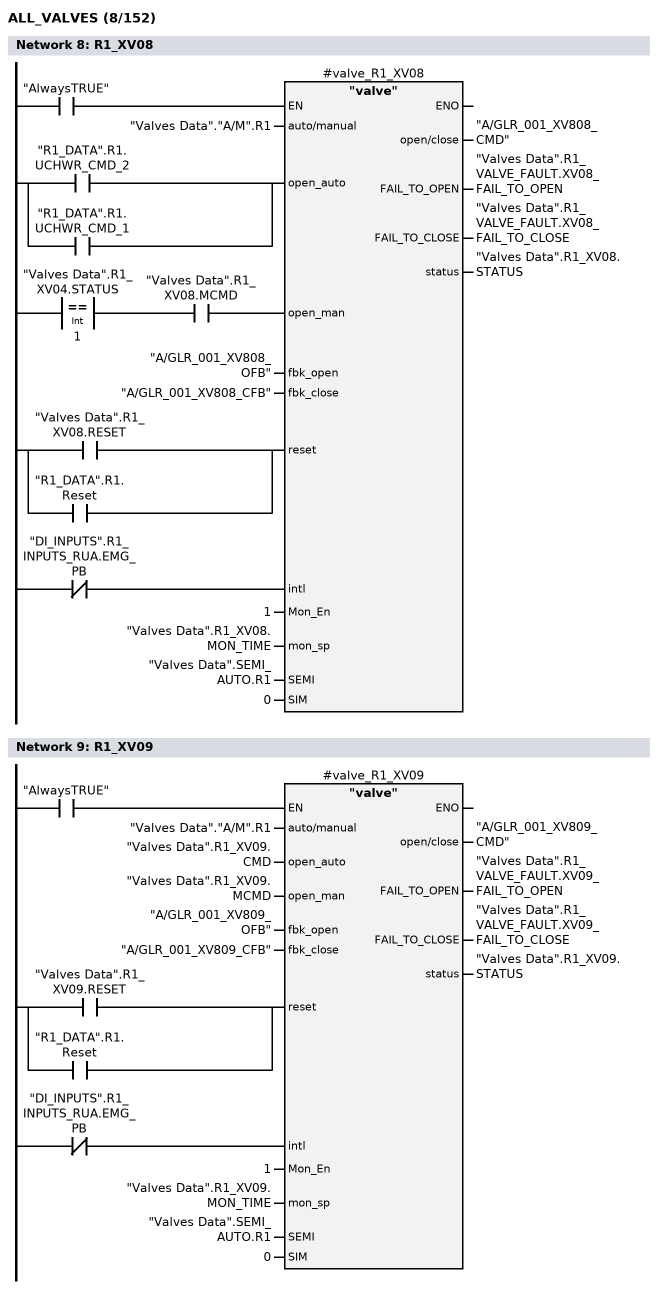
   RUNG wire#powerrail
      Contact( "AlwaysTRUE" )
      #valve_R1_XV08(open_auto := wire#w1, open_man := wire#w2, reset := wire#w3, intl := wire#w4, "auto/manual" := "Valves Data"."A/M".R1, fbk_open := "A/GLR_001_XV808_OFB", fbk_close := "A/GLR_001_XV808_CFB", Mon_En := 1, mon_sp := "Valves Data".R1_XV08.MON_TIME, SEMI := "Valves Data".SEMI_AUTO.R1, SIM := 0, "open/close" => "A/GLR_001_XV808_CMD", FAIL_TO_OPEN => "Valves Data".R1_VALVE_FAULT.XV08_FAIL_TO_OPEN, FAIL_TO_CLOSE => "Valves Data".R1_VALVE_FAULT.XV08_FAIL_TO_CLOSE, status => "Valves Data".R1_XV08.STATUS)
   END_RUNG
   RUNG wire#powerrail
      Contact( "R1_DATA".R1.UCHWR_CMD_2 )
   END_RUNG wire#w1
   RUNG wire#powerrail
      Contact( "R1_DATA".R1.UCHWR_CMD_1 )
   END_RUNG wire#w1
   RUNG wire#powerrail
      { S7_Templates := "SrcType := Int" } EQ_Contact(in1 := "Valves Data".R1_XV04.STATUS, in2 := 1)
      Contact( "Valves Data".R1_XV08.MCMD )
   END_RUNG wire#w2
   RUNG wire#powerrail
      Contact( "Valves Data".R1_XV08.RESET )
   END_RUNG wire#w3
   RUNG wire#powerrail
      Contact( "R1_DATA".R1.Reset )
   END_RUNG wire#w3
   RUNG wire#powerrail
      I_Contact( "DI_INPUTS".R1_INPUTS_RUA.EMG_PB )
   END_RUNG wire#w4
   // the same network as SCL:
   IF "AlwaysTRUE" THEN
       #valve_R1_XV08("auto/manual" := "Valves Data"."A/M".R1,   // "valve"
                      open_auto := "R1_DATA".R1.UCHWR_CMD_2 OR "R1_DATA".R1.UCHWR_CMD_1,
                      open_man := ("Valves Data".R1_XV04.STATUS = 1) AND "Valves Data".R1_XV08.MCMD,
                      fbk_open := "A/GLR_001_XV808_OFB",
                      fbk_close := "A/GLR_001_XV808_CFB",
                      reset := "Valves Data".R1_XV08.RESET OR "R1_DATA".R1.Reset,
                      intl := NOT "DI_INPUTS".R1_INPUTS_RUA.EMG_PB,
                      Mon_En := 1,
                      mon_sp := "Valves Data".R1_XV08.MON_TIME,
                      SEMI := "Valves Data".SEMI_AUTO.R1,
                      SIM := 0,
                      "open/close" => "A/GLR_001_XV808_CMD",
                      FAIL_TO_OPEN => "Valves Data".R1_VALVE_FAULT.XV08_FAIL_TO_OPEN,
                      FAIL_TO_CLOSE => "Valves Data".R1_VALVE_FAULT.XV08_FAIL_TO_CLOSE,
                      status => "Valves Data".R1_XV08.STATUS);
   END_IF;
END_REGION

REGION Network 9: R1_XV09
   RUNG wire#powerrail
      Contact( "AlwaysTRUE" )
      #valve_R1_XV09(reset := wire#w1, intl := wire#w2, "auto/manual" := "Valves Data"."A/M".R1, open_auto := "Valves Data".R1_XV09.CMD, open_man := "Valves Data".R1_XV09.MCMD, fbk_open := "A/GLR_001_XV809_OFB", fbk_close := "A/GLR_001_XV809_CFB", Mon_En := 1, mon_sp := "Valves Data".R1_XV09.MON_TIME, SEMI := "Valves Data".SEMI_AUTO.R1, SIM := 0, "open/close" => "A/GLR_001_XV809_CMD", FAIL_TO_OPEN => "Valves Data".R1_VALVE_FAULT.XV09_FAIL_TO_OPEN, FAIL_TO_CLOSE => "Valves Data".R1_VALVE_FAULT.XV09_FAIL_TO_CLOSE, status => "Valves Data".R1_XV09.STATUS)
   END_RUNG
   RUNG wire#powerrail
      Contact( "Valves Data".R1_XV09.RESET )
   END_RUNG wire#w1
   RUNG wire#powerrail
      Contact( "R1_DATA".R1.Reset )
   END_RUNG wire#w1
   RUNG wire#powerrail
      I_Contact( "DI_INPUTS".R1_INPUTS_RUA.EMG_PB )
   END_RUNG wire#w2
   // the same network as SCL:
   IF "AlwaysTRUE" THEN
       #valve_R1_XV09("auto/manual" := "Valves Data"."A/M".R1,   // "valve"
                      open_auto := "Valves Data".R1_XV09.CMD,
                      open_man := "Valves Data".R1_XV09.MCMD,
                      fbk_open := "A/GLR_001_XV809_OFB",
                      fbk_close := "A/GLR_001_XV809_CFB",
                      reset := "Valves Data".R1_XV09.RESET OR "R1_DATA".R1.Reset,
                      intl := NOT "DI_INPUTS".R1_INPUTS_RUA.EMG_PB,
                      Mon_En := 1,
                      mon_sp := "Valves Data".R1_XV09.MON_TIME,
                      SEMI := "Valves Data".SEMI_AUTO.R1,
                      SIM := 0,
                      "open/close" => "A/GLR_001_XV809_CMD",
                      FAIL_TO_OPEN => "Valves Data".R1_VALVE_FAULT.XV09_FAIL_TO_OPEN,
                      FAIL_TO_CLOSE => "Valves Data".R1_VALVE_FAULT.XV09_FAIL_TO_CLOSE,
                      status => "Valves Data".R1_XV09.STATUS);
   END_IF;
END_REGION

REGION Network 10: R1_XV10
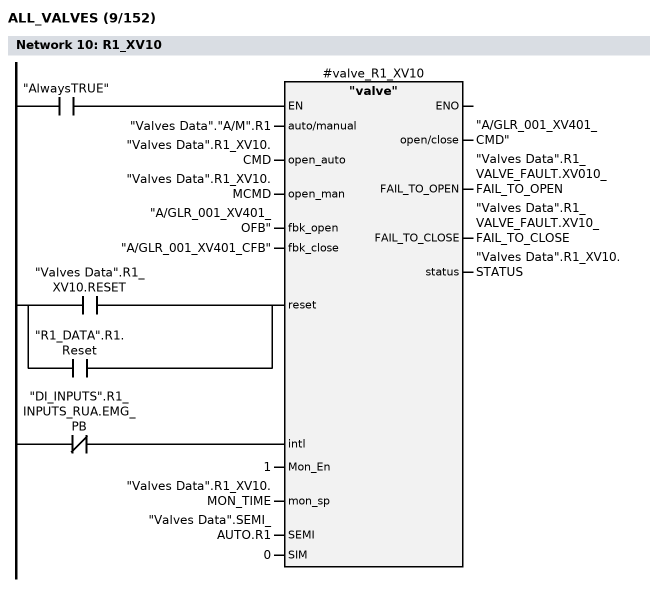
   RUNG wire#powerrail
      Contact( "AlwaysTRUE" )
      #valve_R1_XV10(reset := wire#w1, intl := wire#w2, "auto/manual" := "Valves Data"."A/M".R1, open_auto := "Valves Data".R1_XV10.CMD, open_man := "Valves Data".R1_XV10.MCMD, fbk_open := "A/GLR_001_XV401_OFB", fbk_close := "A/GLR_001_XV401_CFB", Mon_En := 1, mon_sp := "Valves Data".R1_XV10.MON_TIME, SEMI := "Valves Data".SEMI_AUTO.R1, SIM := 0, "open/close" => "A/GLR_001_XV401_CMD", FAIL_TO_OPEN => "Valves Data".R1_VALVE_FAULT.XV010_FAIL_TO_OPEN, FAIL_TO_CLOSE => "Valves Data".R1_VALVE_FAULT.XV10_FAIL_TO_CLOSE, status => "Valves Data".R1_XV10.STATUS)
   END_RUNG
   RUNG wire#powerrail
      Contact( "Valves Data".R1_XV10.RESET )
   END_RUNG wire#w1
   RUNG wire#powerrail
      Contact( "R1_DATA".R1.Reset )
   END_RUNG wire#w1
   RUNG wire#powerrail
      I_Contact( "DI_INPUTS".R1_INPUTS_RUA.EMG_PB )
   END_RUNG wire#w2
   // the same network as SCL:
   IF "AlwaysTRUE" THEN
       #valve_R1_XV10("auto/manual" := "Valves Data"."A/M".R1,   // "valve"
                      open_auto := "Valves Data".R1_XV10.CMD,
                      open_man := "Valves Data".R1_XV10.MCMD,
                      fbk_open := "A/GLR_001_XV401_OFB",
                      fbk_close := "A/GLR_001_XV401_CFB",
                      reset := "Valves Data".R1_XV10.RESET OR "R1_DATA".R1.Reset,
                      intl := NOT "DI_INPUTS".R1_INPUTS_RUA.EMG_PB,
                      Mon_En := 1,
                      mon_sp := "Valves Data".R1_XV10.MON_TIME,
                      SEMI := "Valves Data".SEMI_AUTO.R1,
                      SIM := 0,
                      "open/close" => "A/GLR_001_XV401_CMD",
                      FAIL_TO_OPEN => "Valves Data".R1_VALVE_FAULT.XV010_FAIL_TO_OPEN,
                      FAIL_TO_CLOSE => "Valves Data".R1_VALVE_FAULT.XV10_FAIL_TO_CLOSE,
                      status => "Valves Data".R1_XV10.STATUS);
   END_IF;
END_REGION

REGION Network 11: ****REACTOR_02****
END_REGION

REGION Network 12: R2_XV01
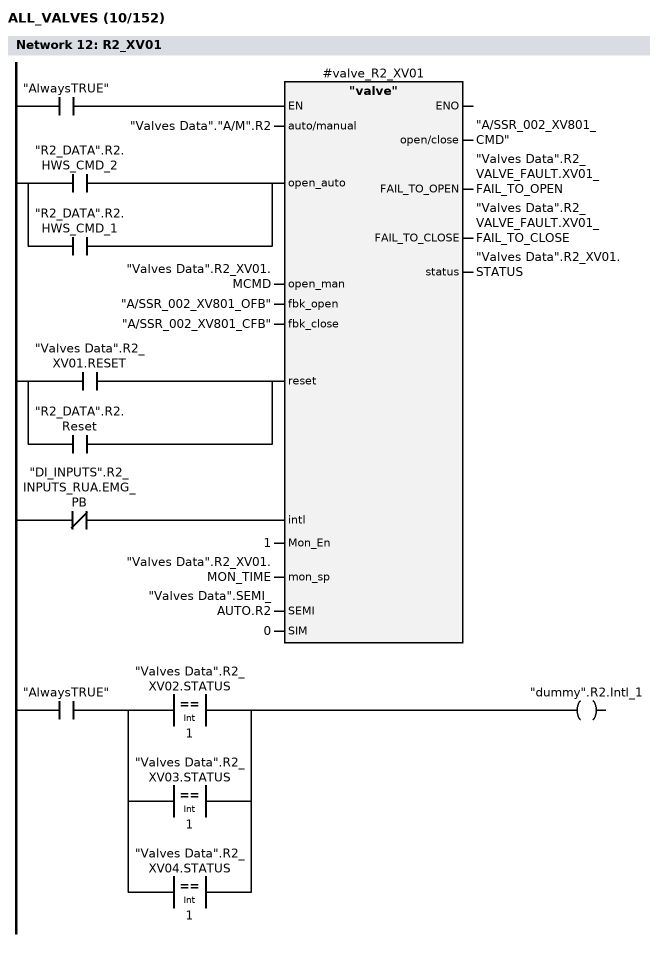
   RUNG wire#powerrail
      Contact( "AlwaysTRUE" )
      #valve_R2_XV01(open_auto := wire#w1, reset := wire#w2, intl := wire#w3, "auto/manual" := "Valves Data"."A/M".R2, open_man := "Valves Data".R2_XV01.MCMD, fbk_open := "A/SSR_002_XV801_OFB", fbk_close := "A/SSR_002_XV801_CFB", Mon_En := 1, mon_sp := "Valves Data".R2_XV01.MON_TIME, SEMI := "Valves Data".SEMI_AUTO.R2, SIM := 0, "open/close" => "A/SSR_002_XV801_CMD", FAIL_TO_OPEN => "Valves Data".R2_VALVE_FAULT.XV01_FAIL_TO_OPEN, FAIL_TO_CLOSE => "Valves Data".R2_VALVE_FAULT.XV01_FAIL_TO_CLOSE, status => "Valves Data".R2_XV01.STATUS)
   END_RUNG
   RUNG wire#powerrail
      Contact( "R2_DATA".R2.HWS_CMD_2 )
   END_RUNG wire#w1
   RUNG wire#powerrail
      Contact( "R2_DATA".R2.HWS_CMD_1 )
   END_RUNG wire#w1
   RUNG wire#powerrail
      Contact( "Valves Data".R2_XV01.RESET )
   END_RUNG wire#w2
   RUNG wire#powerrail
      Contact( "R2_DATA".R2.Reset )
   END_RUNG wire#w2
   RUNG wire#powerrail
      I_Contact( "DI_INPUTS".R2_INPUTS_RUA.EMG_PB )
   END_RUNG wire#w3
   RUNG wire#powerrail
      Contact( "AlwaysTRUE" )
      wire#w4
      { S7_Templates := "SrcType := Int" } EQ_Contact(in1 := "Valves Data".R2_XV02.STATUS, in2 := 1)
      wire#w5
      Coil( "dummy".R2.Intl_1 )
   END_RUNG
   RUNG wire#w4
      { S7_Templates := "SrcType := Int" } EQ_Contact(in1 := "Valves Data".R2_XV03.STATUS, in2 := 1)
   END_RUNG wire#w5
   RUNG wire#w4
      { S7_Templates := "SrcType := Int" } EQ_Contact(in1 := "Valves Data".R2_XV04.STATUS, in2 := 1)
   END_RUNG wire#w5
   // the same network as SCL:
   IF "AlwaysTRUE" THEN
       #valve_R2_XV01("auto/manual" := "Valves Data"."A/M".R2,   // "valve"
                      open_auto := "R2_DATA".R2.HWS_CMD_2 OR "R2_DATA".R2.HWS_CMD_1,
                      open_man := "Valves Data".R2_XV01.MCMD,
                      fbk_open := "A/SSR_002_XV801_OFB",
                      fbk_close := "A/SSR_002_XV801_CFB",
                      reset := "Valves Data".R2_XV01.RESET OR "R2_DATA".R2.Reset,
                      intl := NOT "DI_INPUTS".R2_INPUTS_RUA.EMG_PB,
                      Mon_En := 1,
                      mon_sp := "Valves Data".R2_XV01.MON_TIME,
                      SEMI := "Valves Data".SEMI_AUTO.R2,
                      SIM := 0,
                      "open/close" => "A/SSR_002_XV801_CMD",
                      FAIL_TO_OPEN => "Valves Data".R2_VALVE_FAULT.XV01_FAIL_TO_OPEN,
                      FAIL_TO_CLOSE => "Valves Data".R2_VALVE_FAULT.XV01_FAIL_TO_CLOSE,
                      status => "Valves Data".R2_XV01.STATUS);
   END_IF;
   "dummy".R2.Intl_1 := "AlwaysTRUE" AND (("Valves Data".R2_XV02.STATUS = 1) OR ("Valves Data".R2_XV03.STATUS = 1) OR ("Valves Data".R2_XV04.STATUS = 1));
END_REGION

REGION Network 13: R2_XV02
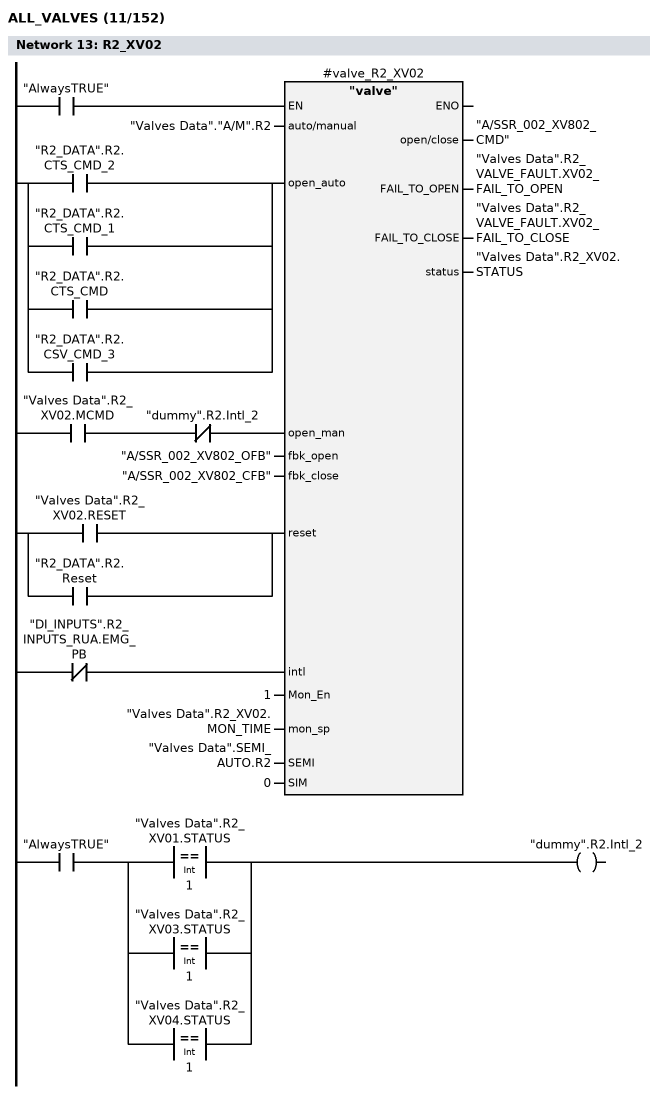
   RUNG wire#powerrail
      Contact( "AlwaysTRUE" )
      #valve_R2_XV02(open_auto := wire#w1, open_man := wire#w2, reset := wire#w3, intl := wire#w4, "auto/manual" := "Valves Data"."A/M".R2, fbk_open := "A/SSR_002_XV802_OFB", fbk_close := "A/SSR_002_XV802_CFB", Mon_En := 1, mon_sp := "Valves Data".R2_XV02.MON_TIME, SEMI := "Valves Data".SEMI_AUTO.R2, SIM := 0, "open/close" => "A/SSR_002_XV802_CMD", FAIL_TO_OPEN => "Valves Data".R2_VALVE_FAULT.XV02_FAIL_TO_OPEN, FAIL_TO_CLOSE => "Valves Data".R2_VALVE_FAULT.XV02_FAIL_TO_CLOSE, status => "Valves Data".R2_XV02.STATUS)
   END_RUNG
   RUNG wire#powerrail
      Contact( "R2_DATA".R2.CTS_CMD_2 )
   END_RUNG wire#w1
   RUNG wire#powerrail
      Contact( "R2_DATA".R2.CTS_CMD_1 )
   END_RUNG wire#w1
   RUNG wire#powerrail
      Contact( "R2_DATA".R2.CTS_CMD )
   END_RUNG wire#w1
   RUNG wire#powerrail
      Contact( "R2_DATA".R2.CSV_CMD_3 )
   END_RUNG wire#w1
   RUNG wire#powerrail
      Contact( "Valves Data".R2_XV02.MCMD )
      I_Contact( "dummy".R2.Intl_2 )
   END_RUNG wire#w2
   RUNG wire#powerrail
      Contact( "Valves Data".R2_XV02.RESET )
   END_RUNG wire#w3
   RUNG wire#powerrail
      Contact( "R2_DATA".R2.Reset )
   END_RUNG wire#w3
   RUNG wire#powerrail
      I_Contact( "DI_INPUTS".R2_INPUTS_RUA.EMG_PB )
   END_RUNG wire#w4
   RUNG wire#powerrail
      Contact( "AlwaysTRUE" )
      wire#w5
      { S7_Templates := "SrcType := Int" } EQ_Contact(in1 := "Valves Data".R2_XV01.STATUS, in2 := 1)
      wire#w6
      Coil( "dummy".R2.Intl_2 )
   END_RUNG
   RUNG wire#w5
      { S7_Templates := "SrcType := Int" } EQ_Contact(in1 := "Valves Data".R2_XV03.STATUS, in2 := 1)
   END_RUNG wire#w6
   RUNG wire#w5
      { S7_Templates := "SrcType := Int" } EQ_Contact(in1 := "Valves Data".R2_XV04.STATUS, in2 := 1)
   END_RUNG wire#w6
   // the same network as SCL:
   IF "AlwaysTRUE" THEN
       #valve_R2_XV02("auto/manual" := "Valves Data"."A/M".R2,   // "valve"
                      open_auto := "R2_DATA".R2.CTS_CMD_2 OR "R2_DATA".R2.CTS_CMD_1 OR "R2_DATA".R2.CTS_CMD OR "R2_DATA".R2.CSV_CMD_3,
                      open_man := "Valves Data".R2_XV02.MCMD AND NOT "dummy".R2.Intl_2,
                      fbk_open := "A/SSR_002_XV802_OFB",
                      fbk_close := "A/SSR_002_XV802_CFB",
                      reset := "Valves Data".R2_XV02.RESET OR "R2_DATA".R2.Reset,
                      intl := NOT "DI_INPUTS".R2_INPUTS_RUA.EMG_PB,
                      Mon_En := 1,
                      mon_sp := "Valves Data".R2_XV02.MON_TIME,
                      SEMI := "Valves Data".SEMI_AUTO.R2,
                      SIM := 0,
                      "open/close" => "A/SSR_002_XV802_CMD",
                      FAIL_TO_OPEN => "Valves Data".R2_VALVE_FAULT.XV02_FAIL_TO_OPEN,
                      FAIL_TO_CLOSE => "Valves Data".R2_VALVE_FAULT.XV02_FAIL_TO_CLOSE,
                      status => "Valves Data".R2_XV02.STATUS);
   END_IF;
   "dummy".R2.Intl_2 := "AlwaysTRUE" AND (("Valves Data".R2_XV01.STATUS = 1) OR ("Valves Data".R2_XV03.STATUS = 1) OR ("Valves Data".R2_XV04.STATUS = 1));
END_REGION

REGION Network 14: R2_XV03
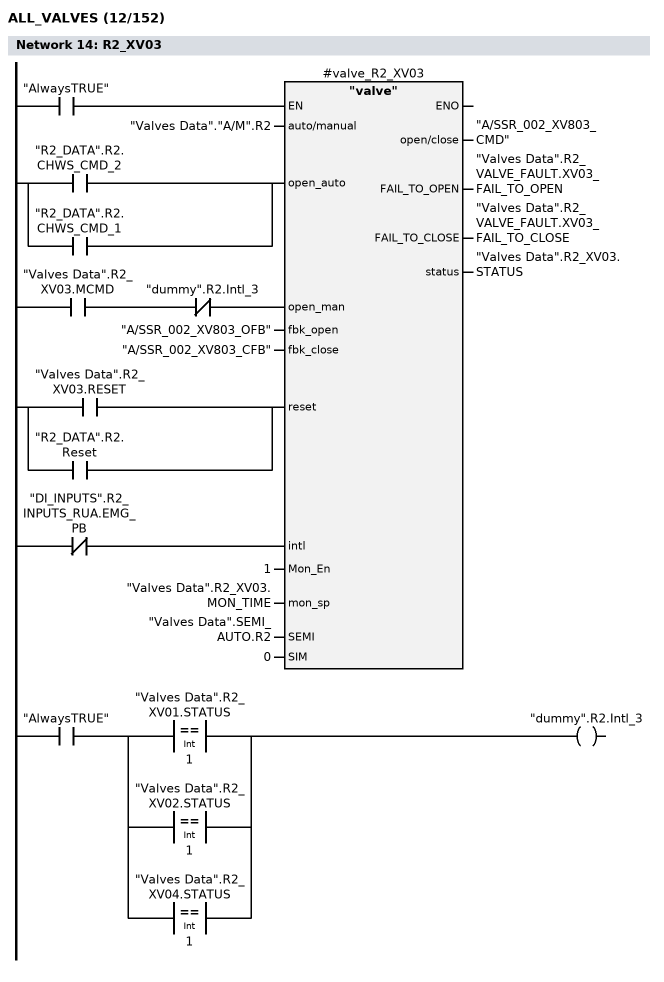
   RUNG wire#powerrail
      Contact( "AlwaysTRUE" )
      #valve_R2_XV03(open_auto := wire#w1, open_man := wire#w2, reset := wire#w3, intl := wire#w4, "auto/manual" := "Valves Data"."A/M".R2, fbk_open := "A/SSR_002_XV803_OFB", fbk_close := "A/SSR_002_XV803_CFB", Mon_En := 1, mon_sp := "Valves Data".R2_XV03.MON_TIME, SEMI := "Valves Data".SEMI_AUTO.R2, SIM := 0, "open/close" => "A/SSR_002_XV803_CMD", FAIL_TO_OPEN => "Valves Data".R2_VALVE_FAULT.XV03_FAIL_TO_OPEN, FAIL_TO_CLOSE => "Valves Data".R2_VALVE_FAULT.XV03_FAIL_TO_CLOSE, status => "Valves Data".R2_XV03.STATUS)
   END_RUNG
   RUNG wire#powerrail
      Contact( "R2_DATA".R2.CHWS_CMD_2 )
   END_RUNG wire#w1
   RUNG wire#powerrail
      Contact( "R2_DATA".R2.CHWS_CMD_1 )
   END_RUNG wire#w1
   RUNG wire#powerrail
      Contact( "Valves Data".R2_XV03.MCMD )
      I_Contact( "dummy".R2.Intl_3 )
   END_RUNG wire#w2
   RUNG wire#powerrail
      Contact( "Valves Data".R2_XV03.RESET )
   END_RUNG wire#w3
   RUNG wire#powerrail
      Contact( "R2_DATA".R2.Reset )
   END_RUNG wire#w3
   RUNG wire#powerrail
      I_Contact( "DI_INPUTS".R2_INPUTS_RUA.EMG_PB )
   END_RUNG wire#w4
   RUNG wire#powerrail
      Contact( "AlwaysTRUE" )
      wire#w5
      { S7_Templates := "SrcType := Int" } EQ_Contact(in1 := "Valves Data".R2_XV01.STATUS, in2 := 1)
      wire#w6
      Coil( "dummy".R2.Intl_3 )
   END_RUNG
   RUNG wire#w5
      { S7_Templates := "SrcType := Int" } EQ_Contact(in1 := "Valves Data".R2_XV02.STATUS, in2 := 1)
   END_RUNG wire#w6
   RUNG wire#w5
      { S7_Templates := "SrcType := Int" } EQ_Contact(in1 := "Valves Data".R2_XV04.STATUS, in2 := 1)
   END_RUNG wire#w6
   // the same network as SCL:
   IF "AlwaysTRUE" THEN
       #valve_R2_XV03("auto/manual" := "Valves Data"."A/M".R2,   // "valve"
                      open_auto := "R2_DATA".R2.CHWS_CMD_2 OR "R2_DATA".R2.CHWS_CMD_1,
                      open_man := "Valves Data".R2_XV03.MCMD AND NOT "dummy".R2.Intl_3,
                      fbk_open := "A/SSR_002_XV803_OFB",
                      fbk_close := "A/SSR_002_XV803_CFB",
                      reset := "Valves Data".R2_XV03.RESET OR "R2_DATA".R2.Reset,
                      intl := NOT "DI_INPUTS".R2_INPUTS_RUA.EMG_PB,
                      Mon_En := 1,
                      mon_sp := "Valves Data".R2_XV03.MON_TIME,
                      SEMI := "Valves Data".SEMI_AUTO.R2,
                      SIM := 0,
                      "open/close" => "A/SSR_002_XV803_CMD",
                      FAIL_TO_OPEN => "Valves Data".R2_VALVE_FAULT.XV03_FAIL_TO_OPEN,
                      FAIL_TO_CLOSE => "Valves Data".R2_VALVE_FAULT.XV03_FAIL_TO_CLOSE,
                      status => "Valves Data".R2_XV03.STATUS);
   END_IF;
   "dummy".R2.Intl_3 := "AlwaysTRUE" AND (("Valves Data".R2_XV01.STATUS = 1) OR ("Valves Data".R2_XV02.STATUS = 1) OR ("Valves Data".R2_XV04.STATUS = 1));
END_REGION

REGION Network 15: R2_XV04
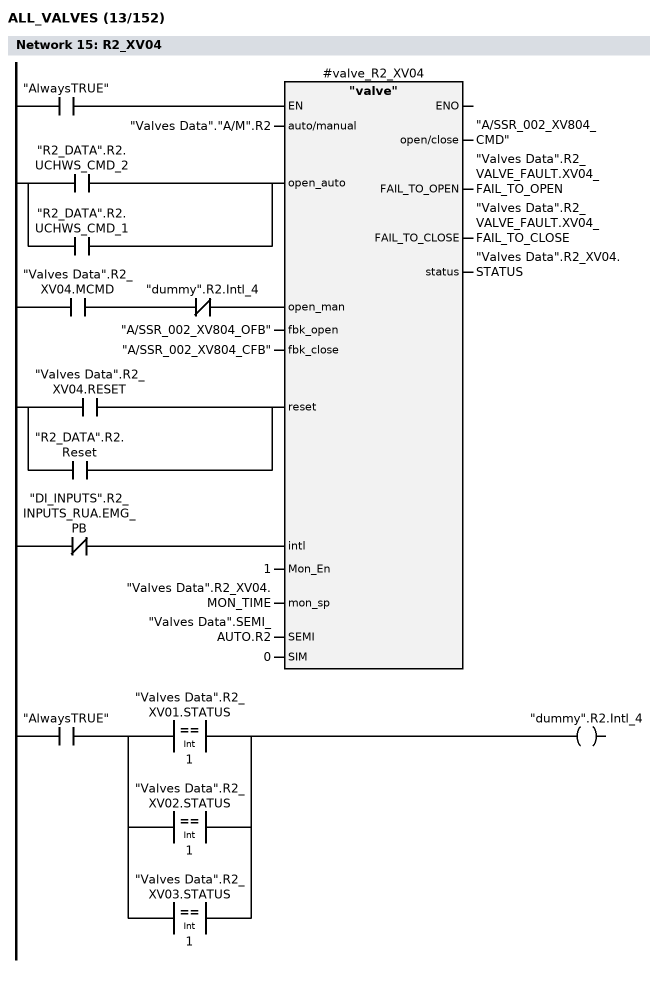
   RUNG wire#powerrail
      Contact( "AlwaysTRUE" )
      #valve_R2_XV04(open_auto := wire#w1, open_man := wire#w2, reset := wire#w3, intl := wire#w4, "auto/manual" := "Valves Data"."A/M".R2, fbk_open := "A/SSR_002_XV804_OFB", fbk_close := "A/SSR_002_XV804_CFB", Mon_En := 1, mon_sp := "Valves Data".R2_XV04.MON_TIME, SEMI := "Valves Data".SEMI_AUTO.R2, SIM := 0, "open/close" => "A/SSR_002_XV804_CMD", FAIL_TO_OPEN => "Valves Data".R2_VALVE_FAULT.XV04_FAIL_TO_OPEN, FAIL_TO_CLOSE => "Valves Data".R2_VALVE_FAULT.XV04_FAIL_TO_CLOSE, status => "Valves Data".R2_XV04.STATUS)
   END_RUNG
   RUNG wire#powerrail
      Contact( "R2_DATA".R2.UCHWS_CMD_2 )
   END_RUNG wire#w1
   RUNG wire#powerrail
      Contact( "R2_DATA".R2.UCHWS_CMD_1 )
   END_RUNG wire#w1
   RUNG wire#powerrail
      Contact( "Valves Data".R2_XV04.MCMD )
      I_Contact( "dummy".R2.Intl_4 )
   END_RUNG wire#w2
   RUNG wire#powerrail
      Contact( "Valves Data".R2_XV04.RESET )
   END_RUNG wire#w3
   RUNG wire#powerrail
      Contact( "R2_DATA".R2.Reset )
   END_RUNG wire#w3
   RUNG wire#powerrail
      I_Contact( "DI_INPUTS".R2_INPUTS_RUA.EMG_PB )
   END_RUNG wire#w4
   RUNG wire#powerrail
      Contact( "AlwaysTRUE" )
      wire#w5
      { S7_Templates := "SrcType := Int" } EQ_Contact(in1 := "Valves Data".R2_XV01.STATUS, in2 := 1)
      wire#w6
      Coil( "dummy".R2.Intl_4 )
   END_RUNG
   RUNG wire#w5
      { S7_Templates := "SrcType := Int" } EQ_Contact(in1 := "Valves Data".R2_XV02.STATUS, in2 := 1)
   END_RUNG wire#w6
   RUNG wire#w5
      { S7_Templates := "SrcType := Int" } EQ_Contact(in1 := "Valves Data".R2_XV03.STATUS, in2 := 1)
   END_RUNG wire#w6
   // the same network as SCL:
   IF "AlwaysTRUE" THEN
       #valve_R2_XV04("auto/manual" := "Valves Data"."A/M".R2,   // "valve"
                      open_auto := "R2_DATA".R2.UCHWS_CMD_2 OR "R2_DATA".R2.UCHWS_CMD_1,
                      open_man := "Valves Data".R2_XV04.MCMD AND NOT "dummy".R2.Intl_4,
                      fbk_open := "A/SSR_002_XV804_OFB",
                      fbk_close := "A/SSR_002_XV804_CFB",
                      reset := "Valves Data".R2_XV04.RESET OR "R2_DATA".R2.Reset,
                      intl := NOT "DI_INPUTS".R2_INPUTS_RUA.EMG_PB,
                      Mon_En := 1,
                      mon_sp := "Valves Data".R2_XV04.MON_TIME,
                      SEMI := "Valves Data".SEMI_AUTO.R2,
                      SIM := 0,
                      "open/close" => "A/SSR_002_XV804_CMD",
                      FAIL_TO_OPEN => "Valves Data".R2_VALVE_FAULT.XV04_FAIL_TO_OPEN,
                      FAIL_TO_CLOSE => "Valves Data".R2_VALVE_FAULT.XV04_FAIL_TO_CLOSE,
                      status => "Valves Data".R2_XV04.STATUS);
   END_IF;
   "dummy".R2.Intl_4 := "AlwaysTRUE" AND (("Valves Data".R2_XV01.STATUS = 1) OR ("Valves Data".R2_XV02.STATUS = 1) OR ("Valves Data".R2_XV03.STATUS = 1));
END_REGION

REGION Network 16: R2_XV05
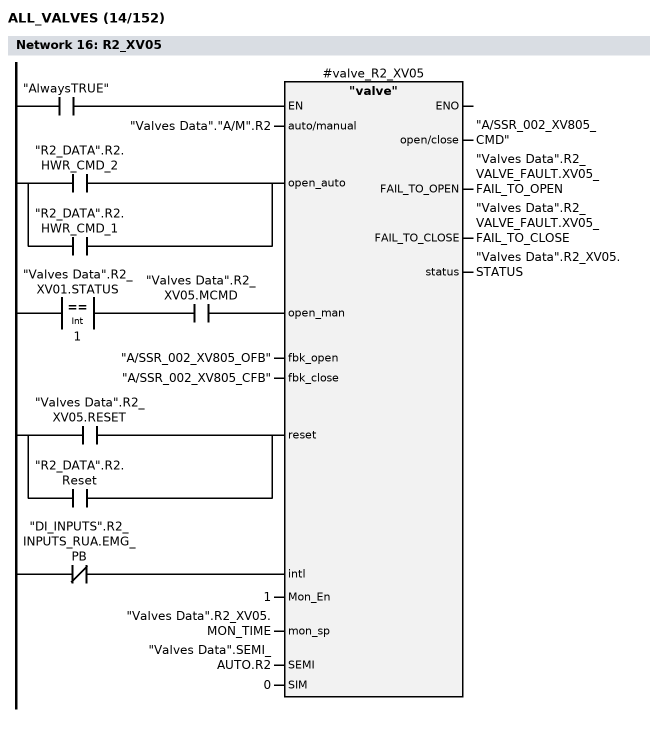
   RUNG wire#powerrail
      Contact( "AlwaysTRUE" )
      #valve_R2_XV05(open_auto := wire#w1, open_man := wire#w2, reset := wire#w3, intl := wire#w4, "auto/manual" := "Valves Data"."A/M".R2, fbk_open := "A/SSR_002_XV805_OFB", fbk_close := "A/SSR_002_XV805_CFB", Mon_En := 1, mon_sp := "Valves Data".R2_XV05.MON_TIME, SEMI := "Valves Data".SEMI_AUTO.R2, SIM := 0, "open/close" => "A/SSR_002_XV805_CMD", FAIL_TO_OPEN => "Valves Data".R2_VALVE_FAULT.XV05_FAIL_TO_OPEN, FAIL_TO_CLOSE => "Valves Data".R2_VALVE_FAULT.XV05_FAIL_TO_CLOSE, status => "Valves Data".R2_XV05.STATUS)
   END_RUNG
   RUNG wire#powerrail
      Contact( "R2_DATA".R2.HWR_CMD_2 )
   END_RUNG wire#w1
   RUNG wire#powerrail
      Contact( "R2_DATA".R2.HWR_CMD_1 )
   END_RUNG wire#w1
   RUNG wire#powerrail
      { S7_Templates := "SrcType := Int" } EQ_Contact(in1 := "Valves Data".R2_XV01.STATUS, in2 := 1)
      Contact( "Valves Data".R2_XV05.MCMD )
   END_RUNG wire#w2
   RUNG wire#powerrail
      Contact( "Valves Data".R2_XV05.RESET )
   END_RUNG wire#w3
   RUNG wire#powerrail
      Contact( "R2_DATA".R2.Reset )
   END_RUNG wire#w3
   RUNG wire#powerrail
      I_Contact( "DI_INPUTS".R2_INPUTS_RUA.EMG_PB )
   END_RUNG wire#w4
   // the same network as SCL:
   IF "AlwaysTRUE" THEN
       #valve_R2_XV05("auto/manual" := "Valves Data"."A/M".R2,   // "valve"
                      open_auto := "R2_DATA".R2.HWR_CMD_2 OR "R2_DATA".R2.HWR_CMD_1,
                      open_man := ("Valves Data".R2_XV01.STATUS = 1) AND "Valves Data".R2_XV05.MCMD,
                      fbk_open := "A/SSR_002_XV805_OFB",
                      fbk_close := "A/SSR_002_XV805_CFB",
                      reset := "Valves Data".R2_XV05.RESET OR "R2_DATA".R2.Reset,
                      intl := NOT "DI_INPUTS".R2_INPUTS_RUA.EMG_PB,
                      Mon_En := 1,
                      mon_sp := "Valves Data".R2_XV05.MON_TIME,
                      SEMI := "Valves Data".SEMI_AUTO.R2,
                      SIM := 0,
                      "open/close" => "A/SSR_002_XV805_CMD",
                      FAIL_TO_OPEN => "Valves Data".R2_VALVE_FAULT.XV05_FAIL_TO_OPEN,
                      FAIL_TO_CLOSE => "Valves Data".R2_VALVE_FAULT.XV05_FAIL_TO_CLOSE,
                      status => "Valves Data".R2_XV05.STATUS);
   END_IF;
END_REGION

REGION Network 17: R2_XV06
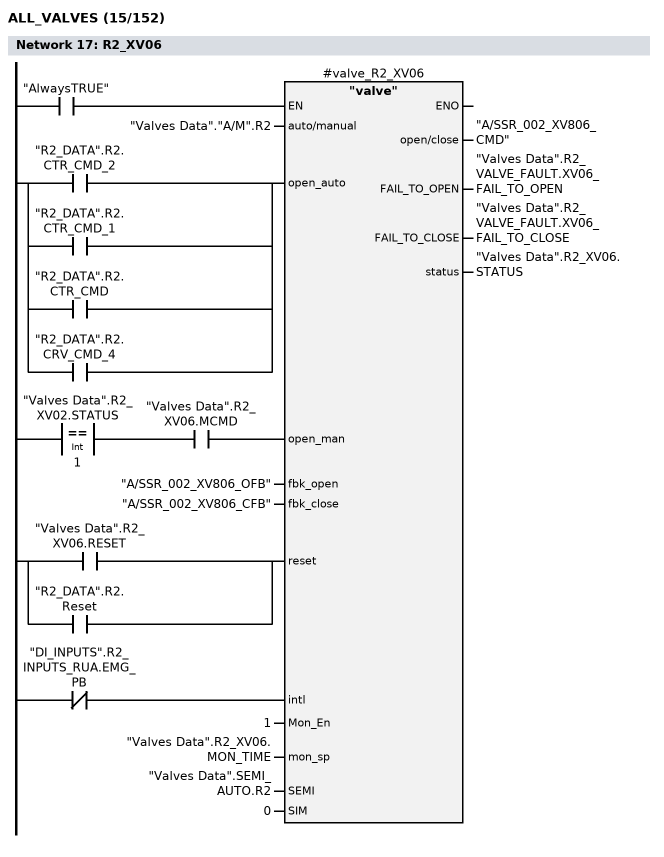
   RUNG wire#powerrail
      Contact( "AlwaysTRUE" )
      #valve_R2_XV06(open_auto := wire#w1, open_man := wire#w2, reset := wire#w3, intl := wire#w4, "auto/manual" := "Valves Data"."A/M".R2, fbk_open := "A/SSR_002_XV806_OFB", fbk_close := "A/SSR_002_XV806_CFB", Mon_En := 1, mon_sp := "Valves Data".R2_XV06.MON_TIME, SEMI := "Valves Data".SEMI_AUTO.R2, SIM := 0, "open/close" => "A/SSR_002_XV806_CMD", FAIL_TO_OPEN => "Valves Data".R2_VALVE_FAULT.XV06_FAIL_TO_OPEN, FAIL_TO_CLOSE => "Valves Data".R2_VALVE_FAULT.XV06_FAIL_TO_CLOSE, status => "Valves Data".R2_XV06.STATUS)
   END_RUNG
   RUNG wire#powerrail
      Contact( "R2_DATA".R2.CTR_CMD_2 )
   END_RUNG wire#w1
   RUNG wire#powerrail
      Contact( "R2_DATA".R2.CTR_CMD_1 )
   END_RUNG wire#w1
   RUNG wire#powerrail
      Contact( "R2_DATA".R2.CTR_CMD )
   END_RUNG wire#w1
   RUNG wire#powerrail
      Contact( "R2_DATA".R2.CRV_CMD_4 )
   END_RUNG wire#w1
   RUNG wire#powerrail
      { S7_Templates := "SrcType := Int" } EQ_Contact(in1 := "Valves Data".R2_XV02.STATUS, in2 := 1)
      Contact( "Valves Data".R2_XV06.MCMD )
   END_RUNG wire#w2
   RUNG wire#powerrail
      Contact( "Valves Data".R2_XV06.RESET )
   END_RUNG wire#w3
   RUNG wire#powerrail
      Contact( "R2_DATA".R2.Reset )
   END_RUNG wire#w3
   RUNG wire#powerrail
      I_Contact( "DI_INPUTS".R2_INPUTS_RUA.EMG_PB )
   END_RUNG wire#w4
   // the same network as SCL:
   IF "AlwaysTRUE" THEN
       #valve_R2_XV06("auto/manual" := "Valves Data"."A/M".R2,   // "valve"
                      open_auto := "R2_DATA".R2.CTR_CMD_2 OR "R2_DATA".R2.CTR_CMD_1 OR "R2_DATA".R2.CTR_CMD OR "R2_DATA".R2.CRV_CMD_4,
                      open_man := ("Valves Data".R2_XV02.STATUS = 1) AND "Valves Data".R2_XV06.MCMD,
                      fbk_open := "A/SSR_002_XV806_OFB",
                      fbk_close := "A/SSR_002_XV806_CFB",
                      reset := "Valves Data".R2_XV06.RESET OR "R2_DATA".R2.Reset,
                      intl := NOT "DI_INPUTS".R2_INPUTS_RUA.EMG_PB,
                      Mon_En := 1,
                      mon_sp := "Valves Data".R2_XV06.MON_TIME,
                      SEMI := "Valves Data".SEMI_AUTO.R2,
                      SIM := 0,
                      "open/close" => "A/SSR_002_XV806_CMD",
                      FAIL_TO_OPEN => "Valves Data".R2_VALVE_FAULT.XV06_FAIL_TO_OPEN,
                      FAIL_TO_CLOSE => "Valves Data".R2_VALVE_FAULT.XV06_FAIL_TO_CLOSE,
                      status => "Valves Data".R2_XV06.STATUS);
   END_IF;
END_REGION

REGION Network 18: R2_XV07
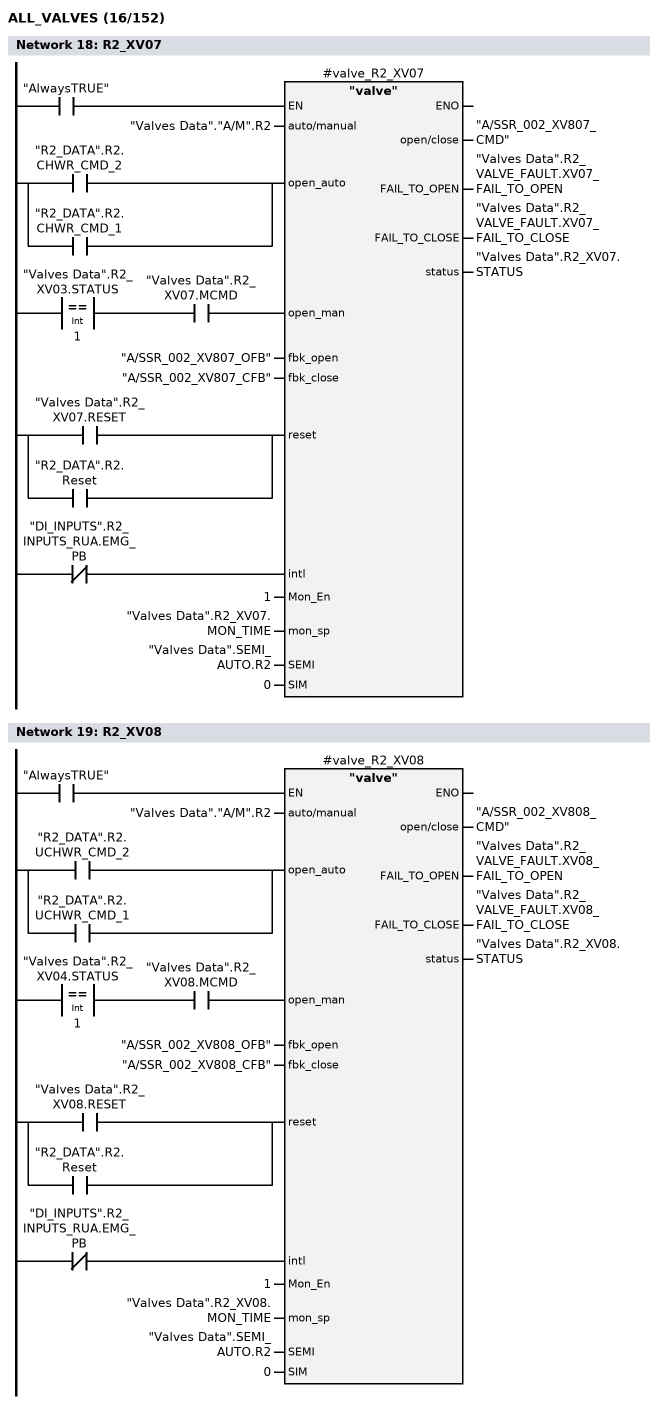
   RUNG wire#powerrail
      Contact( "AlwaysTRUE" )
      #valve_R2_XV07(open_auto := wire#w1, open_man := wire#w2, reset := wire#w3, intl := wire#w4, "auto/manual" := "Valves Data"."A/M".R2, fbk_open := "A/SSR_002_XV807_OFB", fbk_close := "A/SSR_002_XV807_CFB", Mon_En := 1, mon_sp := "Valves Data".R2_XV07.MON_TIME, SEMI := "Valves Data".SEMI_AUTO.R2, SIM := 0, "open/close" => "A/SSR_002_XV807_CMD", FAIL_TO_OPEN => "Valves Data".R2_VALVE_FAULT.XV07_FAIL_TO_OPEN, FAIL_TO_CLOSE => "Valves Data".R2_VALVE_FAULT.XV07_FAIL_TO_CLOSE, status => "Valves Data".R2_XV07.STATUS)
   END_RUNG
   RUNG wire#powerrail
      Contact( "R2_DATA".R2.CHWR_CMD_2 )
   END_RUNG wire#w1
   RUNG wire#powerrail
      Contact( "R2_DATA".R2.CHWR_CMD_1 )
   END_RUNG wire#w1
   RUNG wire#powerrail
      { S7_Templates := "SrcType := Int" } EQ_Contact(in1 := "Valves Data".R2_XV03.STATUS, in2 := 1)
      Contact( "Valves Data".R2_XV07.MCMD )
   END_RUNG wire#w2
   RUNG wire#powerrail
      Contact( "Valves Data".R2_XV07.RESET )
   END_RUNG wire#w3
   RUNG wire#powerrail
      Contact( "R2_DATA".R2.Reset )
   END_RUNG wire#w3
   RUNG wire#powerrail
      I_Contact( "DI_INPUTS".R2_INPUTS_RUA.EMG_PB )
   END_RUNG wire#w4
   // the same network as SCL:
   IF "AlwaysTRUE" THEN
       #valve_R2_XV07("auto/manual" := "Valves Data"."A/M".R2,   // "valve"
                      open_auto := "R2_DATA".R2.CHWR_CMD_2 OR "R2_DATA".R2.CHWR_CMD_1,
                      open_man := ("Valves Data".R2_XV03.STATUS = 1) AND "Valves Data".R2_XV07.MCMD,
                      fbk_open := "A/SSR_002_XV807_OFB",
                      fbk_close := "A/SSR_002_XV807_CFB",
                      reset := "Valves Data".R2_XV07.RESET OR "R2_DATA".R2.Reset,
                      intl := NOT "DI_INPUTS".R2_INPUTS_RUA.EMG_PB,
                      Mon_En := 1,
                      mon_sp := "Valves Data".R2_XV07.MON_TIME,
                      SEMI := "Valves Data".SEMI_AUTO.R2,
                      SIM := 0,
                      "open/close" => "A/SSR_002_XV807_CMD",
                      FAIL_TO_OPEN => "Valves Data".R2_VALVE_FAULT.XV07_FAIL_TO_OPEN,
                      FAIL_TO_CLOSE => "Valves Data".R2_VALVE_FAULT.XV07_FAIL_TO_CLOSE,
                      status => "Valves Data".R2_XV07.STATUS);
   END_IF;
END_REGION

REGION Network 19: R2_XV08
   RUNG wire#powerrail
      Contact( "AlwaysTRUE" )
      #valve_R2_XV08(open_auto := wire#w1, open_man := wire#w2, reset := wire#w3, intl := wire#w4, "auto/manual" := "Valves Data"."A/M".R2, fbk_open := "A/SSR_002_XV808_OFB", fbk_close := "A/SSR_002_XV808_CFB", Mon_En := 1, mon_sp := "Valves Data".R2_XV08.MON_TIME, SEMI := "Valves Data".SEMI_AUTO.R2, SIM := 0, "open/close" => "A/SSR_002_XV808_CMD", FAIL_TO_OPEN => "Valves Data".R2_VALVE_FAULT.XV08_FAIL_TO_OPEN, FAIL_TO_CLOSE => "Valves Data".R2_VALVE_FAULT.XV08_FAIL_TO_CLOSE, status => "Valves Data".R2_XV08.STATUS)
   END_RUNG
   RUNG wire#powerrail
      Contact( "R2_DATA".R2.UCHWR_CMD_2 )
   END_RUNG wire#w1
   RUNG wire#powerrail
      Contact( "R2_DATA".R2.UCHWR_CMD_1 )
   END_RUNG wire#w1
   RUNG wire#powerrail
      { S7_Templates := "SrcType := Int" } EQ_Contact(in1 := "Valves Data".R2_XV04.STATUS, in2 := 1)
      Contact( "Valves Data".R2_XV08.MCMD )
   END_RUNG wire#w2
   RUNG wire#powerrail
      Contact( "Valves Data".R2_XV08.RESET )
   END_RUNG wire#w3
   RUNG wire#powerrail
      Contact( "R2_DATA".R2.Reset )
   END_RUNG wire#w3
   RUNG wire#powerrail
      I_Contact( "DI_INPUTS".R2_INPUTS_RUA.EMG_PB )
   END_RUNG wire#w4
   // the same network as SCL:
   IF "AlwaysTRUE" THEN
       #valve_R2_XV08("auto/manual" := "Valves Data"."A/M".R2,   // "valve"
                      open_auto := "R2_DATA".R2.UCHWR_CMD_2 OR "R2_DATA".R2.UCHWR_CMD_1,
                      open_man := ("Valves Data".R2_XV04.STATUS = 1) AND "Valves Data".R2_XV08.MCMD,
                      fbk_open := "A/SSR_002_XV808_OFB",
                      fbk_close := "A/SSR_002_XV808_CFB",
                      reset := "Valves Data".R2_XV08.RESET OR "R2_DATA".R2.Reset,
                      intl := NOT "DI_INPUTS".R2_INPUTS_RUA.EMG_PB,
                      Mon_En := 1,
                      mon_sp := "Valves Data".R2_XV08.MON_TIME,
                      SEMI := "Valves Data".SEMI_AUTO.R2,
                      SIM := 0,
                      "open/close" => "A/SSR_002_XV808_CMD",
                      FAIL_TO_OPEN => "Valves Data".R2_VALVE_FAULT.XV08_FAIL_TO_OPEN,
                      FAIL_TO_CLOSE => "Valves Data".R2_VALVE_FAULT.XV08_FAIL_TO_CLOSE,
                      status => "Valves Data".R2_XV08.STATUS);
   END_IF;
END_REGION

REGION Network 20: R2_XV09
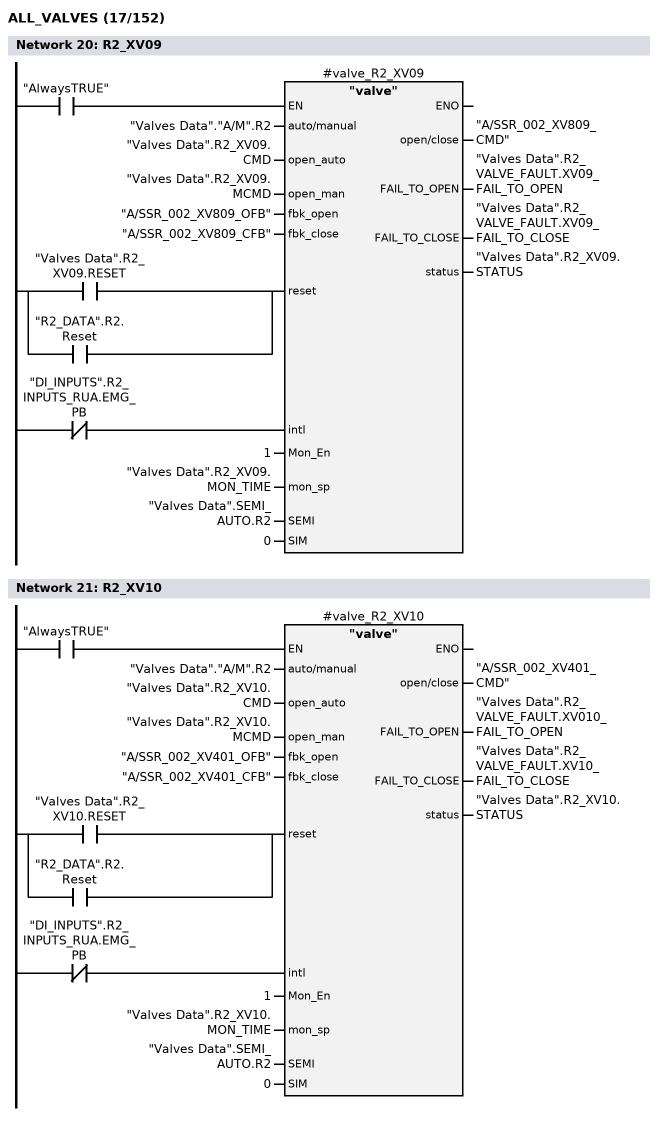
   RUNG wire#powerrail
      Contact( "AlwaysTRUE" )
      #valve_R2_XV09(reset := wire#w1, intl := wire#w2, "auto/manual" := "Valves Data"."A/M".R2, open_auto := "Valves Data".R2_XV09.CMD, open_man := "Valves Data".R2_XV09.MCMD, fbk_open := "A/SSR_002_XV809_OFB", fbk_close := "A/SSR_002_XV809_CFB", Mon_En := 1, mon_sp := "Valves Data".R2_XV09.MON_TIME, SEMI := "Valves Data".SEMI_AUTO.R2, SIM := 0, "open/close" => "A/SSR_002_XV809_CMD", FAIL_TO_OPEN => "Valves Data".R2_VALVE_FAULT.XV09_FAIL_TO_OPEN, FAIL_TO_CLOSE => "Valves Data".R2_VALVE_FAULT.XV09_FAIL_TO_CLOSE, status => "Valves Data".R2_XV09.STATUS)
   END_RUNG
   RUNG wire#powerrail
      Contact( "Valves Data".R2_XV09.RESET )
   END_RUNG wire#w1
   RUNG wire#powerrail
      Contact( "R2_DATA".R2.Reset )
   END_RUNG wire#w1
   RUNG wire#powerrail
      I_Contact( "DI_INPUTS".R2_INPUTS_RUA.EMG_PB )
   END_RUNG wire#w2
   // the same network as SCL:
   IF "AlwaysTRUE" THEN
       #valve_R2_XV09("auto/manual" := "Valves Data"."A/M".R2,   // "valve"
                      open_auto := "Valves Data".R2_XV09.CMD,
                      open_man := "Valves Data".R2_XV09.MCMD,
                      fbk_open := "A/SSR_002_XV809_OFB",
                      fbk_close := "A/SSR_002_XV809_CFB",
                      reset := "Valves Data".R2_XV09.RESET OR "R2_DATA".R2.Reset,
                      intl := NOT "DI_INPUTS".R2_INPUTS_RUA.EMG_PB,
                      Mon_En := 1,
                      mon_sp := "Valves Data".R2_XV09.MON_TIME,
                      SEMI := "Valves Data".SEMI_AUTO.R2,
                      SIM := 0,
                      "open/close" => "A/SSR_002_XV809_CMD",
                      FAIL_TO_OPEN => "Valves Data".R2_VALVE_FAULT.XV09_FAIL_TO_OPEN,
                      FAIL_TO_CLOSE => "Valves Data".R2_VALVE_FAULT.XV09_FAIL_TO_CLOSE,
                      status => "Valves Data".R2_XV09.STATUS);
   END_IF;
END_REGION

REGION Network 21: R2_XV10
   RUNG wire#powerrail
      Contact( "AlwaysTRUE" )
      #valve_R2_XV10(reset := wire#w1, intl := wire#w2, "auto/manual" := "Valves Data"."A/M".R2, open_auto := "Valves Data".R2_XV10.CMD, open_man := "Valves Data".R2_XV10.MCMD, fbk_open := "A/SSR_002_XV401_OFB", fbk_close := "A/SSR_002_XV401_CFB", Mon_En := 1, mon_sp := "Valves Data".R2_XV10.MON_TIME, SEMI := "Valves Data".SEMI_AUTO.R2, SIM := 0, "open/close" => "A/SSR_002_XV401_CMD", FAIL_TO_OPEN => "Valves Data".R2_VALVE_FAULT.XV010_FAIL_TO_OPEN, FAIL_TO_CLOSE => "Valves Data".R2_VALVE_FAULT.XV10_FAIL_TO_CLOSE, status => "Valves Data".R2_XV10.STATUS)
   END_RUNG
   RUNG wire#powerrail
      Contact( "Valves Data".R2_XV10.RESET )
   END_RUNG wire#w1
   RUNG wire#powerrail
      Contact( "R2_DATA".R2.Reset )
   END_RUNG wire#w1
   RUNG wire#powerrail
      I_Contact( "DI_INPUTS".R2_INPUTS_RUA.EMG_PB )
   END_RUNG wire#w2
   // the same network as SCL:
   IF "AlwaysTRUE" THEN
       #valve_R2_XV10("auto/manual" := "Valves Data"."A/M".R2,   // "valve"
                      open_auto := "Valves Data".R2_XV10.CMD,
                      open_man := "Valves Data".R2_XV10.MCMD,
                      fbk_open := "A/SSR_002_XV401_OFB",
                      fbk_close := "A/SSR_002_XV401_CFB",
                      reset := "Valves Data".R2_XV10.RESET OR "R2_DATA".R2.Reset,
                      intl := NOT "DI_INPUTS".R2_INPUTS_RUA.EMG_PB,
                      Mon_En := 1,
                      mon_sp := "Valves Data".R2_XV10.MON_TIME,
                      SEMI := "Valves Data".SEMI_AUTO.R2,
                      SIM := 0,
                      "open/close" => "A/SSR_002_XV401_CMD",
                      FAIL_TO_OPEN => "Valves Data".R2_VALVE_FAULT.XV010_FAIL_TO_OPEN,
                      FAIL_TO_CLOSE => "Valves Data".R2_VALVE_FAULT.XV10_FAIL_TO_CLOSE,
                      status => "Valves Data".R2_XV10.STATUS);
   END_IF;
END_REGION

REGION Network 22: ****REACTOR_03****
END_REGION

REGION Network 23: R3_XV01
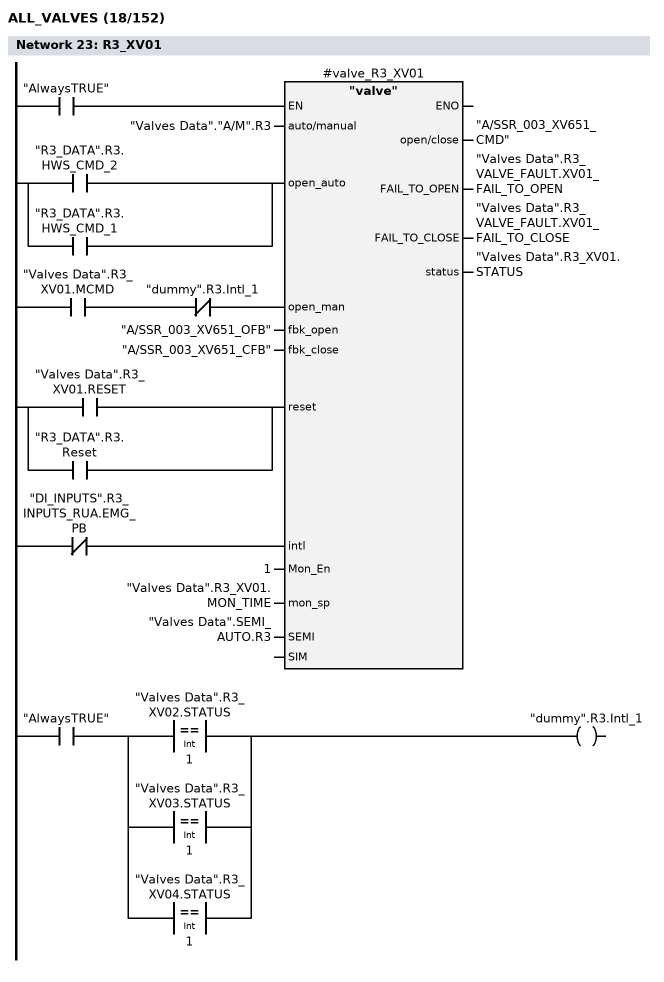
   RUNG wire#powerrail
      Contact( "AlwaysTRUE" )
      #valve_R3_XV01(open_auto := wire#w1, open_man := wire#w2, reset := wire#w3, intl := wire#w4, "auto/manual" := "Valves Data"."A/M".R3, fbk_open := "A/SSR_003_XV651_OFB", fbk_close := "A/SSR_003_XV651_CFB", Mon_En := 1, mon_sp := "Valves Data".R3_XV01.MON_TIME, SEMI := "Valves Data".SEMI_AUTO.R3, SIM :=, "open/close" => "A/SSR_003_XV651_CMD", FAIL_TO_OPEN => "Valves Data".R3_VALVE_FAULT.XV01_FAIL_TO_OPEN, FAIL_TO_CLOSE => "Valves Data".R3_VALVE_FAULT.XV01_FAIL_TO_CLOSE, status => "Valves Data".R3_XV01.STATUS)
   END_RUNG
   RUNG wire#powerrail
      Contact( "R3_DATA".R3.HWS_CMD_2 )
   END_RUNG wire#w1
   RUNG wire#powerrail
      Contact( "R3_DATA".R3.HWS_CMD_1 )
   END_RUNG wire#w1
   RUNG wire#powerrail
      Contact( "Valves Data".R3_XV01.MCMD )
      I_Contact( "dummy".R3.Intl_1 )
   END_RUNG wire#w2
   RUNG wire#powerrail
      Contact( "Valves Data".R3_XV01.RESET )
   END_RUNG wire#w3
   RUNG wire#powerrail
      Contact( "R3_DATA".R3.Reset )
   END_RUNG wire#w3
   RUNG wire#powerrail
      I_Contact( "DI_INPUTS".R3_INPUTS_RUA.EMG_PB )
   END_RUNG wire#w4
   RUNG wire#powerrail
      Contact( "AlwaysTRUE" )
      wire#w5
      { S7_Templates := "SrcType := Int" } EQ_Contact(in1 := "Valves Data".R3_XV02.STATUS, in2 := 1)
      wire#w6
      Coil( "dummy".R3.Intl_1 )
   END_RUNG
   RUNG wire#w5
      { S7_Templates := "SrcType := Int" } EQ_Contact(in1 := "Valves Data".R3_XV03.STATUS, in2 := 1)
   END_RUNG wire#w6
   RUNG wire#w5
      { S7_Templates := "SrcType := Int" } EQ_Contact(in1 := "Valves Data".R3_XV04.STATUS, in2 := 1)
   END_RUNG wire#w6
   // the same network as SCL:
   IF "AlwaysTRUE" THEN
       #valve_R3_XV01("auto/manual" := "Valves Data"."A/M".R3,   // "valve"
                      open_auto := "R3_DATA".R3.HWS_CMD_2 OR "R3_DATA".R3.HWS_CMD_1,
                      open_man := "Valves Data".R3_XV01.MCMD AND NOT "dummy".R3.Intl_1,
                      fbk_open := "A/SSR_003_XV651_OFB",
                      fbk_close := "A/SSR_003_XV651_CFB",
                      reset := "Valves Data".R3_XV01.RESET OR "R3_DATA".R3.Reset,
                      intl := NOT "DI_INPUTS".R3_INPUTS_RUA.EMG_PB,
                      Mon_En := 1,
                      mon_sp := "Valves Data".R3_XV01.MON_TIME,
                      SEMI := "Valves Data".SEMI_AUTO.R3,
                      "open/close" => "A/SSR_003_XV651_CMD",
                      FAIL_TO_OPEN => "Valves Data".R3_VALVE_FAULT.XV01_FAIL_TO_OPEN,
                      FAIL_TO_CLOSE => "Valves Data".R3_VALVE_FAULT.XV01_FAIL_TO_CLOSE,
                      status => "Valves Data".R3_XV01.STATUS);
   END_IF;
   "dummy".R3.Intl_1 := "AlwaysTRUE" AND (("Valves Data".R3_XV02.STATUS = 1) OR ("Valves Data".R3_XV03.STATUS = 1) OR ("Valves Data".R3_XV04.STATUS = 1));
END_REGION

REGION Network 24: R3_XV02
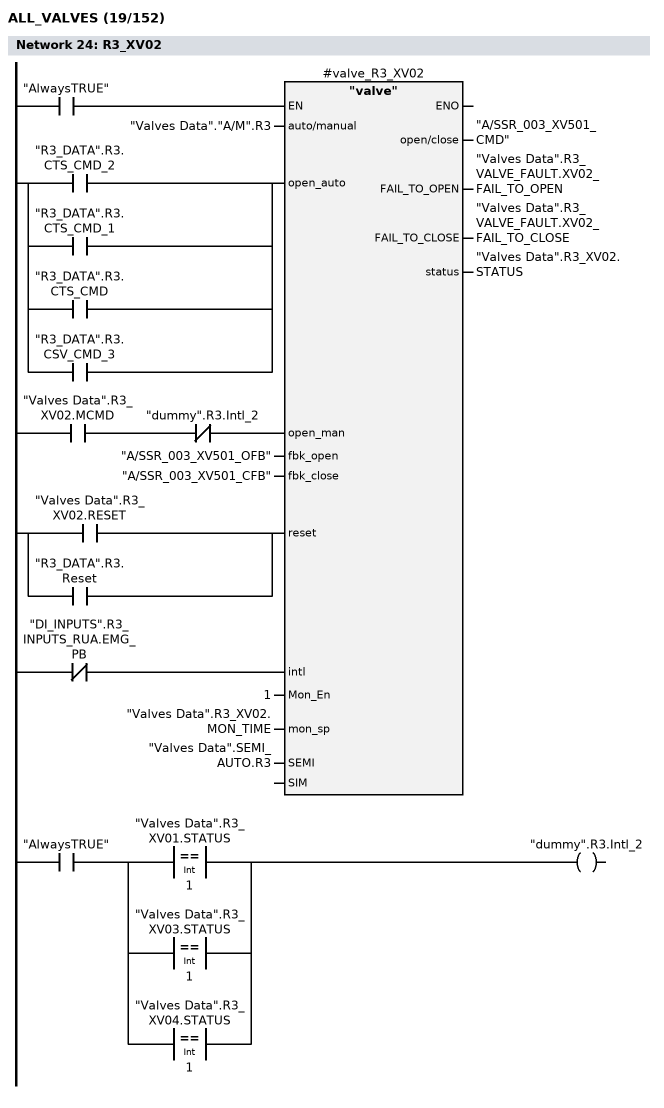
   RUNG wire#powerrail
      Contact( "AlwaysTRUE" )
      #valve_R3_XV02(open_auto := wire#w1, open_man := wire#w2, reset := wire#w3, intl := wire#w4, "auto/manual" := "Valves Data"."A/M".R3, fbk_open := "A/SSR_003_XV501_OFB", fbk_close := "A/SSR_003_XV501_CFB", Mon_En := 1, mon_sp := "Valves Data".R3_XV02.MON_TIME, SEMI := "Valves Data".SEMI_AUTO.R3, SIM :=, "open/close" => "A/SSR_003_XV501_CMD", FAIL_TO_OPEN => "Valves Data".R3_VALVE_FAULT.XV02_FAIL_TO_OPEN, FAIL_TO_CLOSE => "Valves Data".R3_VALVE_FAULT.XV02_FAIL_TO_CLOSE, status => "Valves Data".R3_XV02.STATUS)
   END_RUNG
   RUNG wire#powerrail
      Contact( "R3_DATA".R3.CTS_CMD_2 )
   END_RUNG wire#w1
   RUNG wire#powerrail
      Contact( "R3_DATA".R3.CTS_CMD_1 )
   END_RUNG wire#w1
   RUNG wire#powerrail
      Contact( "R3_DATA".R3.CTS_CMD )
   END_RUNG wire#w1
   RUNG wire#powerrail
      Contact( "R3_DATA".R3.CSV_CMD_3 )
   END_RUNG wire#w1
   RUNG wire#powerrail
      Contact( "Valves Data".R3_XV02.MCMD )
      I_Contact( "dummy".R3.Intl_2 )
   END_RUNG wire#w2
   RUNG wire#powerrail
      Contact( "Valves Data".R3_XV02.RESET )
   END_RUNG wire#w3
   RUNG wire#powerrail
      Contact( "R3_DATA".R3.Reset )
   END_RUNG wire#w3
   RUNG wire#powerrail
      I_Contact( "DI_INPUTS".R3_INPUTS_RUA.EMG_PB )
   END_RUNG wire#w4
   RUNG wire#powerrail
      Contact( "AlwaysTRUE" )
      wire#w5
      { S7_Templates := "SrcType := Int" } EQ_Contact(in1 := "Valves Data".R3_XV01.STATUS, in2 := 1)
      wire#w6
      Coil( "dummy".R3.Intl_2 )
   END_RUNG
   RUNG wire#w5
      { S7_Templates := "SrcType := Int" } EQ_Contact(in1 := "Valves Data".R3_XV03.STATUS, in2 := 1)
   END_RUNG wire#w6
   RUNG wire#w5
      { S7_Templates := "SrcType := Int" } EQ_Contact(in1 := "Valves Data".R3_XV04.STATUS, in2 := 1)
   END_RUNG wire#w6
   // the same network as SCL:
   IF "AlwaysTRUE" THEN
       #valve_R3_XV02("auto/manual" := "Valves Data"."A/M".R3,   // "valve"
                      open_auto := "R3_DATA".R3.CTS_CMD_2 OR "R3_DATA".R3.CTS_CMD_1 OR "R3_DATA".R3.CTS_CMD OR "R3_DATA".R3.CSV_CMD_3,
                      open_man := "Valves Data".R3_XV02.MCMD AND NOT "dummy".R3.Intl_2,
                      fbk_open := "A/SSR_003_XV501_OFB",
                      fbk_close := "A/SSR_003_XV501_CFB",
                      reset := "Valves Data".R3_XV02.RESET OR "R3_DATA".R3.Reset,
                      intl := NOT "DI_INPUTS".R3_INPUTS_RUA.EMG_PB,
                      Mon_En := 1,
                      mon_sp := "Valves Data".R3_XV02.MON_TIME,
                      SEMI := "Valves Data".SEMI_AUTO.R3,
                      "open/close" => "A/SSR_003_XV501_CMD",
                      FAIL_TO_OPEN => "Valves Data".R3_VALVE_FAULT.XV02_FAIL_TO_OPEN,
                      FAIL_TO_CLOSE => "Valves Data".R3_VALVE_FAULT.XV02_FAIL_TO_CLOSE,
                      status => "Valves Data".R3_XV02.STATUS);
   END_IF;
   "dummy".R3.Intl_2 := "AlwaysTRUE" AND (("Valves Data".R3_XV01.STATUS = 1) OR ("Valves Data".R3_XV03.STATUS = 1) OR ("Valves Data".R3_XV04.STATUS = 1));
END_REGION

REGION Network 25: R3_XV03
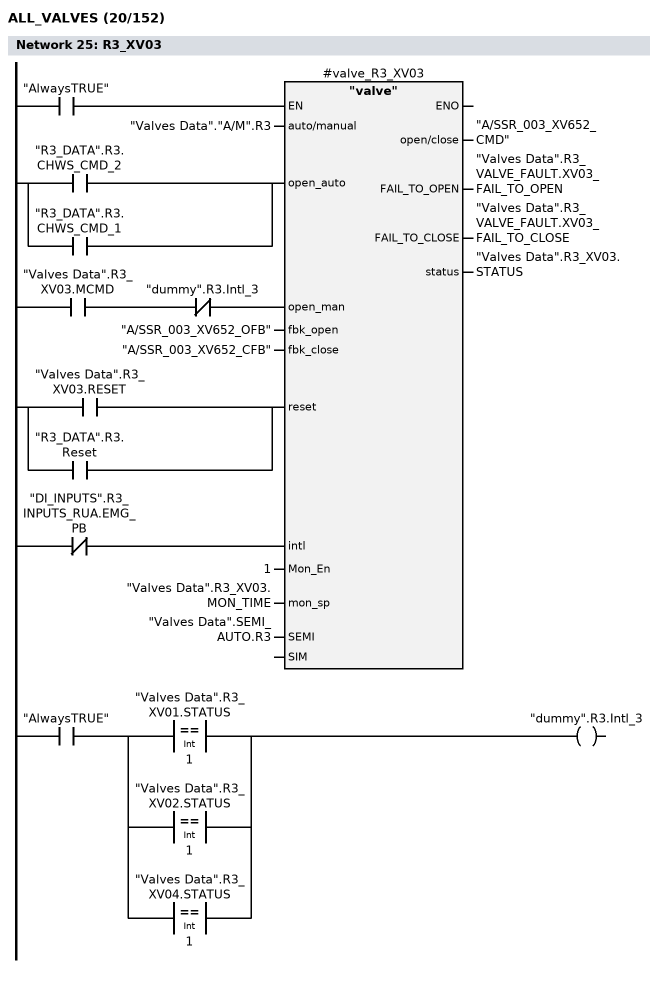
   RUNG wire#powerrail
      Contact( "AlwaysTRUE" )
      #valve_R3_XV03(open_auto := wire#w1, open_man := wire#w2, reset := wire#w3, intl := wire#w4, "auto/manual" := "Valves Data"."A/M".R3, fbk_open := "A/SSR_003_XV652_OFB", fbk_close := "A/SSR_003_XV652_CFB", Mon_En := 1, mon_sp := "Valves Data".R3_XV03.MON_TIME, SEMI := "Valves Data".SEMI_AUTO.R3, SIM :=, "open/close" => "A/SSR_003_XV652_CMD", FAIL_TO_OPEN => "Valves Data".R3_VALVE_FAULT.XV03_FAIL_TO_OPEN, FAIL_TO_CLOSE => "Valves Data".R3_VALVE_FAULT.XV03_FAIL_TO_CLOSE, status => "Valves Data".R3_XV03.STATUS)
   END_RUNG
   RUNG wire#powerrail
      Contact( "R3_DATA".R3.CHWS_CMD_2 )
   END_RUNG wire#w1
   RUNG wire#powerrail
      Contact( "R3_DATA".R3.CHWS_CMD_1 )
   END_RUNG wire#w1
   RUNG wire#powerrail
      Contact( "Valves Data".R3_XV03.MCMD )
      I_Contact( "dummy".R3.Intl_3 )
   END_RUNG wire#w2
   RUNG wire#powerrail
      Contact( "Valves Data".R3_XV03.RESET )
   END_RUNG wire#w3
   RUNG wire#powerrail
      Contact( "R3_DATA".R3.Reset )
   END_RUNG wire#w3
   RUNG wire#powerrail
      I_Contact( "DI_INPUTS".R3_INPUTS_RUA.EMG_PB )
   END_RUNG wire#w4
   RUNG wire#powerrail
      Contact( "AlwaysTRUE" )
      wire#w5
      { S7_Templates := "SrcType := Int" } EQ_Contact(in1 := "Valves Data".R3_XV01.STATUS, in2 := 1)
      wire#w6
      Coil( "dummy".R3.Intl_3 )
   END_RUNG
   RUNG wire#w5
      { S7_Templates := "SrcType := Int" } EQ_Contact(in1 := "Valves Data".R3_XV02.STATUS, in2 := 1)
   END_RUNG wire#w6
   RUNG wire#w5
      { S7_Templates := "SrcType := Int" } EQ_Contact(in1 := "Valves Data".R3_XV04.STATUS, in2 := 1)
   END_RUNG wire#w6
   // the same network as SCL:
   IF "AlwaysTRUE" THEN
       #valve_R3_XV03("auto/manual" := "Valves Data"."A/M".R3,   // "valve"
                      open_auto := "R3_DATA".R3.CHWS_CMD_2 OR "R3_DATA".R3.CHWS_CMD_1,
                      open_man := "Valves Data".R3_XV03.MCMD AND NOT "dummy".R3.Intl_3,
                      fbk_open := "A/SSR_003_XV652_OFB",
                      fbk_close := "A/SSR_003_XV652_CFB",
                      reset := "Valves Data".R3_XV03.RESET OR "R3_DATA".R3.Reset,
                      intl := NOT "DI_INPUTS".R3_INPUTS_RUA.EMG_PB,
                      Mon_En := 1,
                      mon_sp := "Valves Data".R3_XV03.MON_TIME,
                      SEMI := "Valves Data".SEMI_AUTO.R3,
                      "open/close" => "A/SSR_003_XV652_CMD",
                      FAIL_TO_OPEN => "Valves Data".R3_VALVE_FAULT.XV03_FAIL_TO_OPEN,
                      FAIL_TO_CLOSE => "Valves Data".R3_VALVE_FAULT.XV03_FAIL_TO_CLOSE,
                      status => "Valves Data".R3_XV03.STATUS);
   END_IF;
   "dummy".R3.Intl_3 := "AlwaysTRUE" AND (("Valves Data".R3_XV01.STATUS = 1) OR ("Valves Data".R3_XV02.STATUS = 1) OR ("Valves Data".R3_XV04.STATUS = 1));
END_REGION

REGION Network 26: R3_XV04
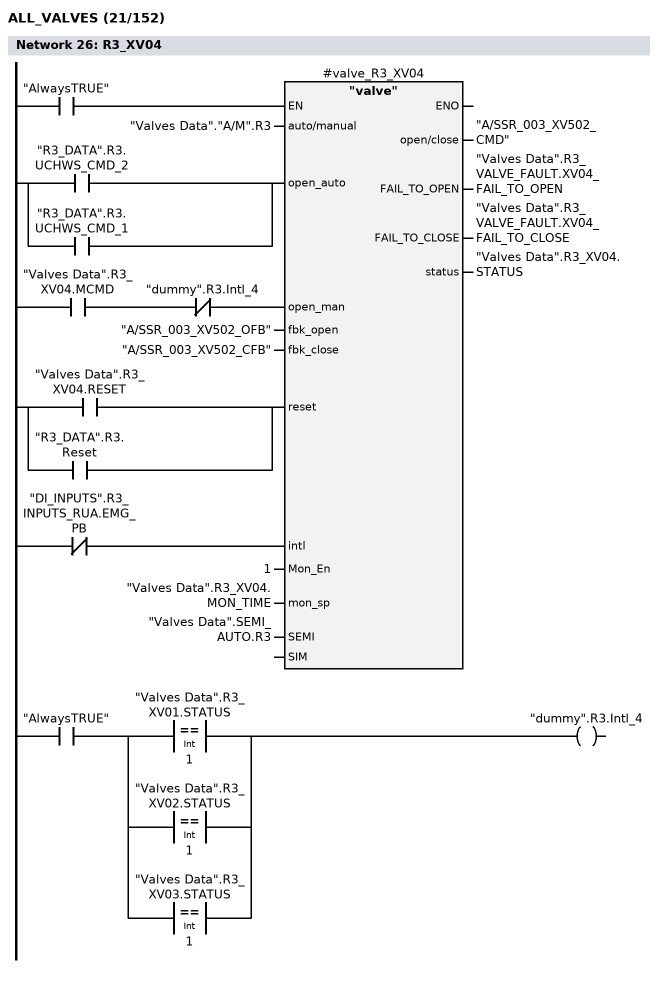
   RUNG wire#powerrail
      Contact( "AlwaysTRUE" )
      #valve_R3_XV04(open_auto := wire#w1, open_man := wire#w2, reset := wire#w3, intl := wire#w4, "auto/manual" := "Valves Data"."A/M".R3, fbk_open := "A/SSR_003_XV502_OFB", fbk_close := "A/SSR_003_XV502_CFB", Mon_En := 1, mon_sp := "Valves Data".R3_XV04.MON_TIME, SEMI := "Valves Data".SEMI_AUTO.R3, SIM :=, "open/close" => "A/SSR_003_XV502_CMD", FAIL_TO_OPEN => "Valves Data".R3_VALVE_FAULT.XV04_FAIL_TO_OPEN, FAIL_TO_CLOSE => "Valves Data".R3_VALVE_FAULT.XV04_FAIL_TO_CLOSE, status => "Valves Data".R3_XV04.STATUS)
   END_RUNG
   RUNG wire#powerrail
      Contact( "R3_DATA".R3.UCHWS_CMD_2 )
   END_RUNG wire#w1
   RUNG wire#powerrail
      Contact( "R3_DATA".R3.UCHWS_CMD_1 )
   END_RUNG wire#w1
   RUNG wire#powerrail
      Contact( "Valves Data".R3_XV04.MCMD )
      I_Contact( "dummy".R3.Intl_4 )
   END_RUNG wire#w2
   RUNG wire#powerrail
      Contact( "Valves Data".R3_XV04.RESET )
   END_RUNG wire#w3
   RUNG wire#powerrail
      Contact( "R3_DATA".R3.Reset )
   END_RUNG wire#w3
   RUNG wire#powerrail
      I_Contact( "DI_INPUTS".R3_INPUTS_RUA.EMG_PB )
   END_RUNG wire#w4
   RUNG wire#powerrail
      Contact( "AlwaysTRUE" )
      wire#w5
      { S7_Templates := "SrcType := Int" } EQ_Contact(in1 := "Valves Data".R3_XV01.STATUS, in2 := 1)
      wire#w6
      Coil( "dummy".R3.Intl_4 )
   END_RUNG
   RUNG wire#w5
      { S7_Templates := "SrcType := Int" } EQ_Contact(in1 := "Valves Data".R3_XV02.STATUS, in2 := 1)
   END_RUNG wire#w6
   RUNG wire#w5
      { S7_Templates := "SrcType := Int" } EQ_Contact(in1 := "Valves Data".R3_XV03.STATUS, in2 := 1)
   END_RUNG wire#w6
   // the same network as SCL:
   IF "AlwaysTRUE" THEN
       #valve_R3_XV04("auto/manual" := "Valves Data"."A/M".R3,   // "valve"
                      open_auto := "R3_DATA".R3.UCHWS_CMD_2 OR "R3_DATA".R3.UCHWS_CMD_1,
                      open_man := "Valves Data".R3_XV04.MCMD AND NOT "dummy".R3.Intl_4,
                      fbk_open := "A/SSR_003_XV502_OFB",
                      fbk_close := "A/SSR_003_XV502_CFB",
                      reset := "Valves Data".R3_XV04.RESET OR "R3_DATA".R3.Reset,
                      intl := NOT "DI_INPUTS".R3_INPUTS_RUA.EMG_PB,
                      Mon_En := 1,
                      mon_sp := "Valves Data".R3_XV04.MON_TIME,
                      SEMI := "Valves Data".SEMI_AUTO.R3,
                      "open/close" => "A/SSR_003_XV502_CMD",
                      FAIL_TO_OPEN => "Valves Data".R3_VALVE_FAULT.XV04_FAIL_TO_OPEN,
                      FAIL_TO_CLOSE => "Valves Data".R3_VALVE_FAULT.XV04_FAIL_TO_CLOSE,
                      status => "Valves Data".R3_XV04.STATUS);
   END_IF;
   "dummy".R3.Intl_4 := "AlwaysTRUE" AND (("Valves Data".R3_XV01.STATUS = 1) OR ("Valves Data".R3_XV02.STATUS = 1) OR ("Valves Data".R3_XV03.STATUS = 1));
END_REGION

REGION Network 27: R3_XV05
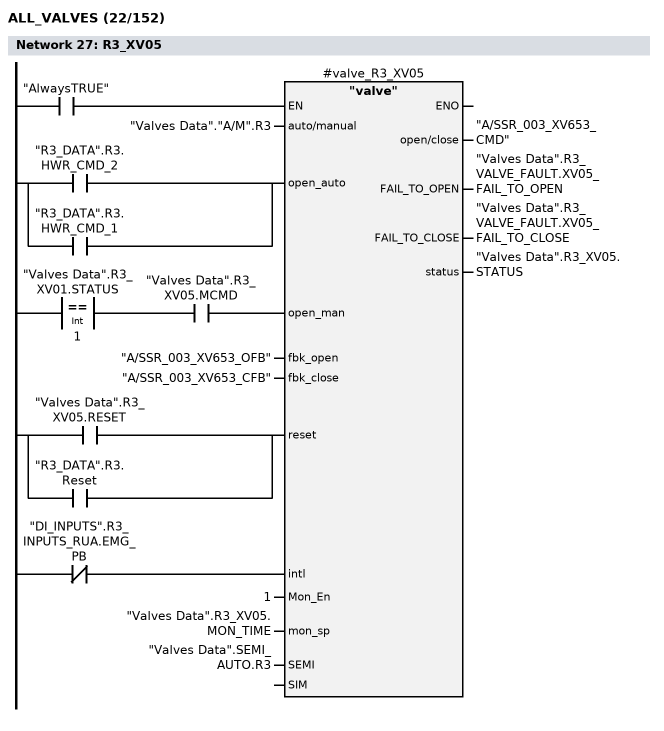
   RUNG wire#powerrail
      Contact( "AlwaysTRUE" )
      #valve_R3_XV05(open_auto := wire#w1, open_man := wire#w2, reset := wire#w3, intl := wire#w4, "auto/manual" := "Valves Data"."A/M".R3, fbk_open := "A/SSR_003_XV653_OFB", fbk_close := "A/SSR_003_XV653_CFB", Mon_En := 1, mon_sp := "Valves Data".R3_XV05.MON_TIME, SEMI := "Valves Data".SEMI_AUTO.R3, SIM :=, "open/close" => "A/SSR_003_XV653_CMD", FAIL_TO_OPEN => "Valves Data".R3_VALVE_FAULT.XV05_FAIL_TO_OPEN, FAIL_TO_CLOSE => "Valves Data".R3_VALVE_FAULT.XV05_FAIL_TO_CLOSE, status => "Valves Data".R3_XV05.STATUS)
   END_RUNG
   RUNG wire#powerrail
      Contact( "R3_DATA".R3.HWR_CMD_2 )
   END_RUNG wire#w1
   RUNG wire#powerrail
      Contact( "R3_DATA".R3.HWR_CMD_1 )
   END_RUNG wire#w1
   RUNG wire#powerrail
      { S7_Templates := "SrcType := Int" } EQ_Contact(in1 := "Valves Data".R3_XV01.STATUS, in2 := 1)
      Contact( "Valves Data".R3_XV05.MCMD )
   END_RUNG wire#w2
   RUNG wire#powerrail
      Contact( "Valves Data".R3_XV05.RESET )
   END_RUNG wire#w3
   RUNG wire#powerrail
      Contact( "R3_DATA".R3.Reset )
   END_RUNG wire#w3
   RUNG wire#powerrail
      I_Contact( "DI_INPUTS".R3_INPUTS_RUA.EMG_PB )
   END_RUNG wire#w4
   // the same network as SCL:
   IF "AlwaysTRUE" THEN
       #valve_R3_XV05("auto/manual" := "Valves Data"."A/M".R3,   // "valve"
                      open_auto := "R3_DATA".R3.HWR_CMD_2 OR "R3_DATA".R3.HWR_CMD_1,
                      open_man := ("Valves Data".R3_XV01.STATUS = 1) AND "Valves Data".R3_XV05.MCMD,
                      fbk_open := "A/SSR_003_XV653_OFB",
                      fbk_close := "A/SSR_003_XV653_CFB",
                      reset := "Valves Data".R3_XV05.RESET OR "R3_DATA".R3.Reset,
                      intl := NOT "DI_INPUTS".R3_INPUTS_RUA.EMG_PB,
                      Mon_En := 1,
                      mon_sp := "Valves Data".R3_XV05.MON_TIME,
                      SEMI := "Valves Data".SEMI_AUTO.R3,
                      "open/close" => "A/SSR_003_XV653_CMD",
                      FAIL_TO_OPEN => "Valves Data".R3_VALVE_FAULT.XV05_FAIL_TO_OPEN,
                      FAIL_TO_CLOSE => "Valves Data".R3_VALVE_FAULT.XV05_FAIL_TO_CLOSE,
                      status => "Valves Data".R3_XV05.STATUS);
   END_IF;
END_REGION

REGION Network 28: R3_XV06
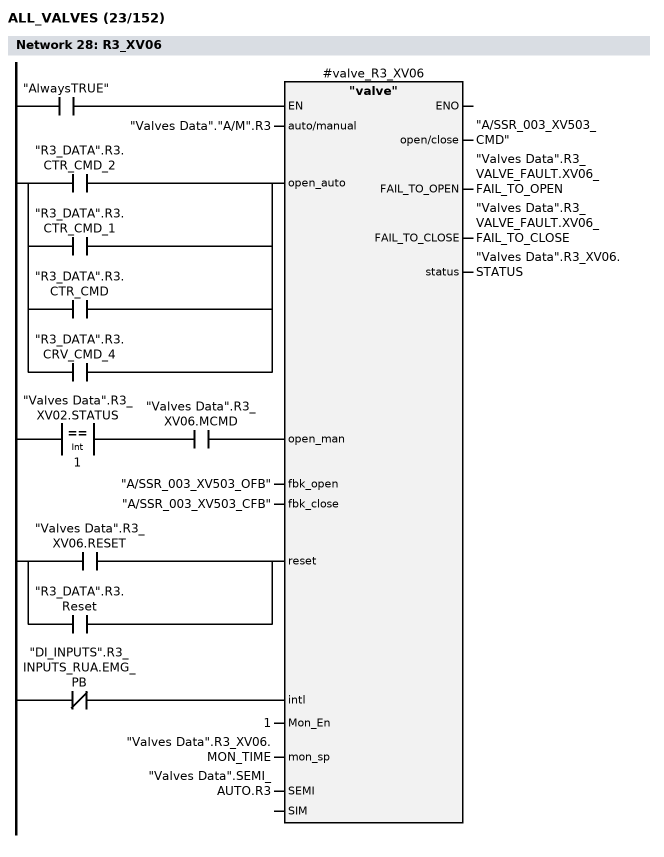
   RUNG wire#powerrail
      Contact( "AlwaysTRUE" )
      #valve_R3_XV06(open_auto := wire#w1, open_man := wire#w2, reset := wire#w3, intl := wire#w4, "auto/manual" := "Valves Data"."A/M".R3, fbk_open := "A/SSR_003_XV503_OFB", fbk_close := "A/SSR_003_XV503_CFB", Mon_En := 1, mon_sp := "Valves Data".R3_XV06.MON_TIME, SEMI := "Valves Data".SEMI_AUTO.R3, SIM :=, "open/close" => "A/SSR_003_XV503_CMD", FAIL_TO_OPEN => "Valves Data".R3_VALVE_FAULT.XV06_FAIL_TO_OPEN, FAIL_TO_CLOSE => "Valves Data".R3_VALVE_FAULT.XV06_FAIL_TO_CLOSE, status => "Valves Data".R3_XV06.STATUS)
   END_RUNG
   RUNG wire#powerrail
      Contact( "R3_DATA".R3.CTR_CMD_2 )
   END_RUNG wire#w1
   RUNG wire#powerrail
      Contact( "R3_DATA".R3.CTR_CMD_1 )
   END_RUNG wire#w1
   RUNG wire#powerrail
      Contact( "R3_DATA".R3.CTR_CMD )
   END_RUNG wire#w1
   RUNG wire#powerrail
      Contact( "R3_DATA".R3.CRV_CMD_4 )
   END_RUNG wire#w1
   RUNG wire#powerrail
      { S7_Templates := "SrcType := Int" } EQ_Contact(in1 := "Valves Data".R3_XV02.STATUS, in2 := 1)
      Contact( "Valves Data".R3_XV06.MCMD )
   END_RUNG wire#w2
   RUNG wire#powerrail
      Contact( "Valves Data".R3_XV06.RESET )
   END_RUNG wire#w3
   RUNG wire#powerrail
      Contact( "R3_DATA".R3.Reset )
   END_RUNG wire#w3
   RUNG wire#powerrail
      I_Contact( "DI_INPUTS".R3_INPUTS_RUA.EMG_PB )
   END_RUNG wire#w4
   // the same network as SCL:
   IF "AlwaysTRUE" THEN
       #valve_R3_XV06("auto/manual" := "Valves Data"."A/M".R3,   // "valve"
                      open_auto := "R3_DATA".R3.CTR_CMD_2 OR "R3_DATA".R3.CTR_CMD_1 OR "R3_DATA".R3.CTR_CMD OR "R3_DATA".R3.CRV_CMD_4,
                      open_man := ("Valves Data".R3_XV02.STATUS = 1) AND "Valves Data".R3_XV06.MCMD,
                      fbk_open := "A/SSR_003_XV503_OFB",
                      fbk_close := "A/SSR_003_XV503_CFB",
                      reset := "Valves Data".R3_XV06.RESET OR "R3_DATA".R3.Reset,
                      intl := NOT "DI_INPUTS".R3_INPUTS_RUA.EMG_PB,
                      Mon_En := 1,
                      mon_sp := "Valves Data".R3_XV06.MON_TIME,
                      SEMI := "Valves Data".SEMI_AUTO.R3,
                      "open/close" => "A/SSR_003_XV503_CMD",
                      FAIL_TO_OPEN => "Valves Data".R3_VALVE_FAULT.XV06_FAIL_TO_OPEN,
                      FAIL_TO_CLOSE => "Valves Data".R3_VALVE_FAULT.XV06_FAIL_TO_CLOSE,
                      status => "Valves Data".R3_XV06.STATUS);
   END_IF;
END_REGION

REGION Network 29: R3_XV07
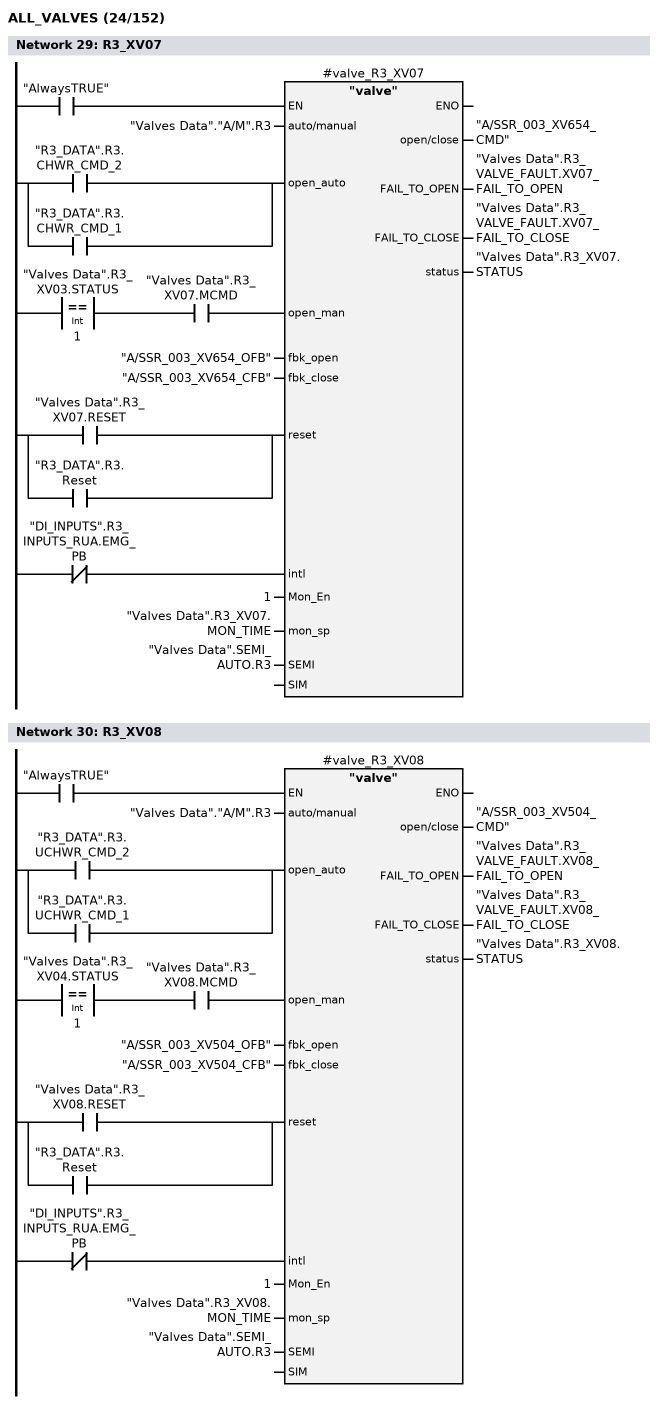
   RUNG wire#powerrail
      Contact( "AlwaysTRUE" )
      #valve_R3_XV07(open_auto := wire#w1, open_man := wire#w2, reset := wire#w3, intl := wire#w4, "auto/manual" := "Valves Data"."A/M".R3, fbk_open := "A/SSR_003_XV654_OFB", fbk_close := "A/SSR_003_XV654_CFB", Mon_En := 1, mon_sp := "Valves Data".R3_XV07.MON_TIME, SEMI := "Valves Data".SEMI_AUTO.R3, SIM :=, "open/close" => "A/SSR_003_XV654_CMD", FAIL_TO_OPEN => "Valves Data".R3_VALVE_FAULT.XV07_FAIL_TO_OPEN, FAIL_TO_CLOSE => "Valves Data".R3_VALVE_FAULT.XV07_FAIL_TO_CLOSE, status => "Valves Data".R3_XV07.STATUS)
   END_RUNG
   RUNG wire#powerrail
      Contact( "R3_DATA".R3.CHWR_CMD_2 )
   END_RUNG wire#w1
   RUNG wire#powerrail
      Contact( "R3_DATA".R3.CHWR_CMD_1 )
   END_RUNG wire#w1
   RUNG wire#powerrail
      { S7_Templates := "SrcType := Int" } EQ_Contact(in1 := "Valves Data".R3_XV03.STATUS, in2 := 1)
      Contact( "Valves Data".R3_XV07.MCMD )
   END_RUNG wire#w2
   RUNG wire#powerrail
      Contact( "Valves Data".R3_XV07.RESET )
   END_RUNG wire#w3
   RUNG wire#powerrail
      Contact( "R3_DATA".R3.Reset )
   END_RUNG wire#w3
   RUNG wire#powerrail
      I_Contact( "DI_INPUTS".R3_INPUTS_RUA.EMG_PB )
   END_RUNG wire#w4
   // the same network as SCL:
   IF "AlwaysTRUE" THEN
       #valve_R3_XV07("auto/manual" := "Valves Data"."A/M".R3,   // "valve"
                      open_auto := "R3_DATA".R3.CHWR_CMD_2 OR "R3_DATA".R3.CHWR_CMD_1,
                      open_man := ("Valves Data".R3_XV03.STATUS = 1) AND "Valves Data".R3_XV07.MCMD,
                      fbk_open := "A/SSR_003_XV654_OFB",
                      fbk_close := "A/SSR_003_XV654_CFB",
                      reset := "Valves Data".R3_XV07.RESET OR "R3_DATA".R3.Reset,
                      intl := NOT "DI_INPUTS".R3_INPUTS_RUA.EMG_PB,
                      Mon_En := 1,
                      mon_sp := "Valves Data".R3_XV07.MON_TIME,
                      SEMI := "Valves Data".SEMI_AUTO.R3,
                      "open/close" => "A/SSR_003_XV654_CMD",
                      FAIL_TO_OPEN => "Valves Data".R3_VALVE_FAULT.XV07_FAIL_TO_OPEN,
                      FAIL_TO_CLOSE => "Valves Data".R3_VALVE_FAULT.XV07_FAIL_TO_CLOSE,
                      status => "Valves Data".R3_XV07.STATUS);
   END_IF;
END_REGION

REGION Network 30: R3_XV08
   RUNG wire#powerrail
      Contact( "AlwaysTRUE" )
      #valve_R3_XV08(open_auto := wire#w1, open_man := wire#w2, reset := wire#w3, intl := wire#w4, "auto/manual" := "Valves Data"."A/M".R3, fbk_open := "A/SSR_003_XV504_OFB", fbk_close := "A/SSR_003_XV504_CFB", Mon_En := 1, mon_sp := "Valves Data".R3_XV08.MON_TIME, SEMI := "Valves Data".SEMI_AUTO.R3, SIM :=, "open/close" => "A/SSR_003_XV504_CMD", FAIL_TO_OPEN => "Valves Data".R3_VALVE_FAULT.XV08_FAIL_TO_OPEN, FAIL_TO_CLOSE => "Valves Data".R3_VALVE_FAULT.XV08_FAIL_TO_CLOSE, status => "Valves Data".R3_XV08.STATUS)
   END_RUNG
   RUNG wire#powerrail
      Contact( "R3_DATA".R3.UCHWR_CMD_2 )
   END_RUNG wire#w1
   RUNG wire#powerrail
      Contact( "R3_DATA".R3.UCHWR_CMD_1 )
   END_RUNG wire#w1
   RUNG wire#powerrail
      { S7_Templates := "SrcType := Int" } EQ_Contact(in1 := "Valves Data".R3_XV04.STATUS, in2 := 1)
      Contact( "Valves Data".R3_XV08.MCMD )
   END_RUNG wire#w2
   RUNG wire#powerrail
      Contact( "Valves Data".R3_XV08.RESET )
   END_RUNG wire#w3
   RUNG wire#powerrail
      Contact( "R3_DATA".R3.Reset )
   END_RUNG wire#w3
   RUNG wire#powerrail
      I_Contact( "DI_INPUTS".R3_INPUTS_RUA.EMG_PB )
   END_RUNG wire#w4
   // the same network as SCL:
   IF "AlwaysTRUE" THEN
       #valve_R3_XV08("auto/manual" := "Valves Data"."A/M".R3,   // "valve"
                      open_auto := "R3_DATA".R3.UCHWR_CMD_2 OR "R3_DATA".R3.UCHWR_CMD_1,
                      open_man := ("Valves Data".R3_XV04.STATUS = 1) AND "Valves Data".R3_XV08.MCMD,
                      fbk_open := "A/SSR_003_XV504_OFB",
                      fbk_close := "A/SSR_003_XV504_CFB",
                      reset := "Valves Data".R3_XV08.RESET OR "R3_DATA".R3.Reset,
                      intl := NOT "DI_INPUTS".R3_INPUTS_RUA.EMG_PB,
                      Mon_En := 1,
                      mon_sp := "Valves Data".R3_XV08.MON_TIME,
                      SEMI := "Valves Data".SEMI_AUTO.R3,
                      "open/close" => "A/SSR_003_XV504_CMD",
                      FAIL_TO_OPEN => "Valves Data".R3_VALVE_FAULT.XV08_FAIL_TO_OPEN,
                      FAIL_TO_CLOSE => "Valves Data".R3_VALVE_FAULT.XV08_FAIL_TO_CLOSE,
                      status => "Valves Data".R3_XV08.STATUS);
   END_IF;
END_REGION

REGION Network 31: R3_XV09
